(* IEC 61131-3 sources: trust-platform/examples/room_heating/libraries/plant/src, 22 files *)

(* ---- types.st ---- *)
(* The Plant library's shared types (specification trust-plant-library §3–§9). *)
NAMESPACE Plant

(* Who commands a device (§3): the program in Auto, the operator in Manual. *)
TYPE E_Mode : (Auto, Manual, OutOfService); END_TYPE

(* A measurement's quality (§7.1). *)
TYPE E_Quality : (Good, Uncertain, Bad); END_TYPE

(* A sequence's state (§9.4). *)
TYPE E_SequenceState : (Idle, Running, Held, Stopping, Stopped, Completed, Aborted, Failed); END_TYPE

END_NAMESPACE

(* ---- interfaces.st ---- *)
(* The capabilities of the Plant blocks (specification trust-plant-library §5). Each interface is
   small; a block implements the ones it supports. Operator commands return TRUE when accepted.
   An HMI button may call only a method of an interface its block implements. *)
NAMESPACE Plant

(* Mode and reset, common to every device (§3). *)
INTERFACE IDevice
    METHOD SetMode : BOOL
    VAR_INPUT
        Value : E_Mode;
    END_VAR
    END_METHOD
    METHOD GetMode : E_Mode
    END_METHOD
    METHOD Reset : BOOL
    END_METHOD
END_INTERFACE

INTERFACE IRunDevice EXTENDS IDevice
    METHOD Start : BOOL
    END_METHOD
    METHOD Stop : BOOL
    END_METHOD
    METHOD IsRunning : BOOL
    END_METHOD
END_INTERFACE

INTERFACE ISpeedDevice EXTENDS IRunDevice
    METHOD SetSpeed : BOOL
    VAR_INPUT
        Value : LREAL;
    END_VAR
    END_METHOD
END_INTERFACE

INTERFACE IPowerDevice EXTENDS IRunDevice
    METHOD SetPower : BOOL
    VAR_INPUT
        Value : LREAL;
    END_VAR
    END_METHOD
END_INTERFACE

INTERFACE IReversingDevice EXTENDS IDevice
    METHOD StartForward : BOOL
    END_METHOD
    METHOD StartReverse : BOOL
    END_METHOD
    METHOD Stop : BOOL
    END_METHOD
END_INTERFACE

INTERFACE ITwoSpeedDevice EXTENDS IDevice
    METHOD StartSlow : BOOL
    END_METHOD
    METHOD StartFast : BOOL
    END_METHOD
    METHOD Stop : BOOL
    END_METHOD
END_INTERFACE

INTERFACE IOpenCloseDevice EXTENDS IDevice
    METHOD Open : BOOL
    END_METHOD
    METHOD Close : BOOL
    END_METHOD
    METHOD IsOpen : BOOL
    END_METHOD
    METHOD IsClosed : BOOL
    END_METHOD
END_INTERFACE

(* A motor-operated valve can stop between its end positions. *)
INTERFACE ITravelStop
    METHOD StopTravel : BOOL
    END_METHOD
END_INTERFACE

INTERFACE IExtendRetractDevice EXTENDS IDevice
    METHOD Extend : BOOL
    END_METHOD
    METHOD Retract : BOOL
    END_METHOD
    METHOD IsExtended : BOOL
    END_METHOD
    METHOD IsRetracted : BOOL
    END_METHOD
END_INTERFACE

INTERFACE IPositionDevice EXTENDS IDevice
    METHOD SetPosition : BOOL
    VAR_INPUT
        Value : LREAL;
    END_VAR
    END_METHOD
    METHOD GetPosition : LREAL
    END_METHOD
END_INTERFACE

(* A device that a controller drives through its Auto value (§5): FollowsAuto is TRUE while the
   device follows that value now, GetActualValue is what the device does. A loop tracks
   GetActualValue while FollowsAuto is FALSE (§8.1), so it neither winds up nor bumps when the
   device follows it again. *)
INTERFACE IControlledDevice
    METHOD FollowsAuto : BOOL
    END_METHOD
    METHOD GetActualValue : LREAL
    END_METHOD
END_INTERFACE

(* An Engineer confirms that the service is done (§4.7). *)
INTERFACE IServiceable
    METHOD ServiceDone : BOOL
    END_METHOD
END_INTERFACE

(* A run device a group can command in Auto (§9.2). *)
INTERFACE IDutyMember EXTENDS IRunDevice
    METHOD IsAvailable : BOOL
    END_METHOD
    METHOD Demand
    VAR_INPUT
        Run : BOOL;
    END_VAR
    END_METHOD
    METHOD GetRunHours : LREAL
    END_METHOD
END_INTERFACE

INTERFACE IMeasurement
    METHOD GetValue : LREAL
    END_METHOD
    METHOD GetQuality : E_Quality
    END_METHOD
END_INTERFACE

INTERFACE ITotal
    METHOD ResetTotal : BOOL
    END_METHOD
END_INTERFACE

INTERFACE ICounter
    METHOD ResetCount : BOOL
    END_METHOD
END_INTERFACE

INTERFACE ITare
    METHOD Tare : BOOL
    END_METHOD
    METHOD ClearTare : BOOL
    END_METHOD
END_INTERFACE

INTERFACE ISetpoint
    METHOD SetSetpoint : BOOL
    VAR_INPUT
        Value : LREAL;
    END_VAR
    END_METHOD
END_INTERFACE

(* An Engineer bypasses one condition of a set for a limited time (§9.1). *)
INTERFACE IBypass
    METHOD Bypass : BOOL
    VAR_INPUT
        Index : INT;
    END_VAR
    END_METHOD
    METHOD RemoveBypass : BOOL
    VAR_INPUT
        Index : INT;
    END_VAR
    END_METHOD
END_INTERFACE

(* The alarms a block holds, for an alarm manager (§4.5, §9.3). *)
INTERFACE IAlarmSource
    METHOD GetAlarmCount : INT
    END_METHOD
    METHOD GetAlarm : REF_TO Alarm.Alarm
    VAR_INPUT
        Index : INT;
    END_VAR
    END_METHOD
END_INTERFACE

INTERFACE IAlarmManager
    METHOD AcknowledgeAll : BOOL
    END_METHOD
    METHOD Silence : BOOL
    END_METHOD
END_INTERFACE

INTERFACE ISequence
    METHOD Start : BOOL
    END_METHOD
    METHOD Stop : BOOL
    END_METHOD
    METHOD Hold : BOOL
    END_METHOD
    METHOD Resume : BOOL
    END_METHOD
    METHOD Abort : BOOL
    END_METHOD
    METHOD Reset : BOOL
    END_METHOD
    METHOD GetState : E_SequenceState
    END_METHOD
END_INTERFACE

INTERFACE ISequenceManager
    METHOD StopAll : BOOL
    END_METHOD
    METHOD AbortAll : BOOL
    END_METHOD
END_INTERFACE

END_NAMESPACE

(* ---- analog_input.st ---- *)
(* Analog instruments (specification trust-plant-library §7.1): scaling, quality, the optional
   Control.LowPass filter and four limit alarms. A broken signal raises one signal alarm and
   suppresses the limit alarms. The defaults suit a 4-20 mA signal (NAMUR NE 43); set RawLow,
   RawHigh, BadBelow and BadAbove for other signals. *)
NAMESPACE Plant
USING Alarm;
USING Control;

FUNCTION_BLOCK FB_AnalogInput IMPLEMENTS IMeasurement, IAlarmSource
VAR_INPUT
    (* The channel's value, for example in mA. *)
    Raw : LREAL;
    (* The I/O module's diagnosis for this channel. *)
    SignalFault : BOOL;
END_VAR
VAR PUBLIC
    Unit : STRING[16];
END_VAR
VAR PUBLIC RETAIN
    RawLow : LREAL := 4.0;
    RawHigh : LREAL := 20.0;
    RangeLow : LREAL := 0.0;
    RangeHigh : LREAL := 100.0;
    BadBelow : LREAL := 3.6;
    BadAbove : LREAL := 21.0;
    FilterTime : TIME := T#0s;
    HighHighEnabled : BOOL;
    HighEnabled : BOOL;
    LowEnabled : BOOL;
    LowLowEnabled : BOOL;
    HighHighLimit : LREAL := 95.0;
    HighLimit : LREAL := 90.0;
    LowLimit : LREAL := 10.0;
    LowLowLimit : LREAL := 5.0;
    Deadband : LREAL := 1.0;
    AlarmDelay : TIME := T#0s;
END_VAR
VAR_OUTPUT NON_RETAIN
    Value : LREAL;
    Percent : LREAL;
    Quality : E_Quality := E_Quality#Bad;
    Fault : BOOL;
    HighHigh : BOOL;
    High : BOOL;
    Low : BOOL;
    LowLow : BOOL;
END_VAR
VAR NON_RETAIN
    Filter : LowPass;
    Filtering : BOOL;
    HasValue : BOOL;
    Clock : FB_ScanClock;
    SignalAlarm : Alarm.DigitalAlarm;
    HighHighAlarm : Alarm.LimitAlarm;
    HighAlarm : Alarm.LimitAlarm;
    LowAlarm : Alarm.LimitAlarm;
    LowLowAlarm : Alarm.LimitAlarm;
END_VAR
    Measure();

METHOD PROTECTED Measure
VAR
    Span : LREAL;
    Range : LREAL;
    Scaled : LREAL;
    Parameters : LowPassParameters;
END_VAR
    Clock();
    Span := RawHigh - RawLow;
    Range := RangeHigh - RangeLow;
    IF NOT SignalFault AND F_Finite(Raw) AND Raw >= BadBelow AND Raw <= BadAbove
        AND F_Finite(Span) AND Span <> 0.0 THEN
        Scaled := RangeLow + (Raw - RawLow) * Range / Span;
        IF FilterTime > T#0s AND HasValue THEN
            Parameters.TimeConstant := F_Seconds(FilterTime);
            Parameters.Order := FilterOrder#FirstOrder;
            Filter.Configure(Parameters := Parameters);
            IF NOT Filtering THEN
                Filter.Initialize(Input := Value);
                Filtering := TRUE;
            END_IF;
            IF Clock.Seconds > 0.0 THEN
                Value := Filter.Update(Input := Scaled, CycleTime := Clock.Seconds);
            END_IF;
        ELSE
            Value := Scaled;
            Filtering := FALSE;
        END_IF;
        HasValue := TRUE;
        Quality := E_Quality#Good;
    ELSE
        (* The value holds its last good reading. *)
        Quality := E_Quality#Bad;
        Filtering := FALSE;
    END_IF;
    Fault := Quality = E_Quality#Bad;
    IF Range <> 0.0 AND F_Finite(Range) THEN
        Percent := (Value - RangeLow) / Range * 100.0;
    ELSE
        Percent := 0.0;
    END_IF;

    (* A limit that is not enabled, and every limit while the signal is bad, is suppressed: it
       does not annunciate and its output stays FALSE. *)
    SignalAlarm(Condition := Fault, Message := 'Signal fault', Priority := AlarmPriority#Medium);
    HighHighAlarm(Value := Value, Limit := HighHighLimit, Deadband := ABS(Deadband),
        Direction := LimitDirection#High, OnDelay := AlarmDelay, Suppressed := Fault OR NOT HighHighEnabled,
        Message := 'High-high', Priority := AlarmPriority#High);
    HighAlarm(Value := Value, Limit := HighLimit, Deadband := ABS(Deadband),
        Direction := LimitDirection#High, OnDelay := AlarmDelay, Suppressed := Fault OR NOT HighEnabled,
        Message := 'High', Priority := AlarmPriority#Medium);
    LowAlarm(Value := Value, Limit := LowLimit, Deadband := ABS(Deadband),
        Direction := LimitDirection#Low, OnDelay := AlarmDelay, Suppressed := Fault OR NOT LowEnabled,
        Message := 'Low', Priority := AlarmPriority#Medium);
    LowLowAlarm(Value := Value, Limit := LowLowLimit, Deadband := ABS(Deadband),
        Direction := LimitDirection#Low, OnDelay := AlarmDelay, Suppressed := Fault OR NOT LowLowEnabled,
        Message := 'Low-low', Priority := AlarmPriority#High);
    HighHigh := HighHighAlarm.Active AND NOT HighHighAlarm.SuppressedByDesign;
    High := HighAlarm.Active AND NOT HighAlarm.SuppressedByDesign;
    Low := LowAlarm.Active AND NOT LowAlarm.SuppressedByDesign;
    LowLow := LowLowAlarm.Active AND NOT LowLowAlarm.SuppressedByDesign;
END_METHOD

METHOD PUBLIC GetValue : LREAL
    GetValue := Value;
END_METHOD

METHOD PUBLIC GetQuality : E_Quality
    GetQuality := Quality;
END_METHOD

METHOD PUBLIC GetAlarmCount : INT
    GetAlarmCount := 5;
END_METHOD

METHOD PUBLIC GetAlarm : REF_TO Alarm.Alarm
VAR_INPUT
    Index : INT;
END_VAR
    CASE Index OF
        1: GetAlarm := REF(SignalAlarm);
        2: GetAlarm := REF(HighHighAlarm);
        3: GetAlarm := REF(HighAlarm);
        4: GetAlarm := REF(LowAlarm);
        5: GetAlarm := REF(LowLowAlarm);
    ELSE
        GetAlarm := NULL;
    END_CASE;
END_METHOD
END_FUNCTION_BLOCK

(* The instruments below differ in name and symbol; their unit comes from the instance. *)
FUNCTION_BLOCK FB_LevelInput EXTENDS FB_AnalogInput
    Measure();
END_FUNCTION_BLOCK

FUNCTION_BLOCK FB_PressureInput EXTENDS FB_AnalogInput
    Measure();
END_FUNCTION_BLOCK

FUNCTION_BLOCK FB_TemperatureInput EXTENDS FB_AnalogInput
    Measure();
END_FUNCTION_BLOCK

FUNCTION_BLOCK FB_AnalyzerInput EXTENDS FB_AnalogInput
    Measure();
END_FUNCTION_BLOCK

(* A flow instrument with its own totaliser on its measured value (§7.1.6). *)
FUNCTION_BLOCK FB_FlowInput EXTENDS FB_AnalogInput IMPLEMENTS ITotal
VAR_OUTPUT RETAIN
    (* Retained as well as the totaliser's, so it reads right before the first scan. *)
    Total : LREAL;
END_VAR
VAR PUBLIC RETAIN
    (* The time base of the flow's unit: T#1h for m3/h. *)
    TotalPer : TIME := T#1h;
END_VAR
VAR
    Totalizer : FB_Totalizer;
END_VAR
    Measure();
    Totalizer.TotalPer := TotalPer;
    Totalizer(Rate := Value, RateGood := Quality = E_Quality#Good);
    Total := Totalizer.Total;

METHOD PUBLIC ResetTotal : BOOL
    ResetTotal := Totalizer.ResetTotal();
    Total := 0.0;
END_METHOD
END_FUNCTION_BLOCK

END_NAMESPACE

(* ---- conditions.st ---- *)
(* Condition sets (specification trust-plant-library §9.1): up to eight conditions with texts, a
   first-out text, and Engineer bypasses that end by themselves. Interlocks and permissives may
   be bypassed; protection may not. These are ordinary process conditions, not certified safety
   functions. *)
NAMESPACE Plant

FUNCTION_BLOCK ABSTRACT FB_ConditionSet
VAR_INPUT
    (* TRUE while the condition is healthy; an unused condition stays TRUE. *)
    Condition1 : BOOL := TRUE;
    Condition2 : BOOL := TRUE;
    Condition3 : BOOL := TRUE;
    Condition4 : BOOL := TRUE;
    Condition5 : BOOL := TRUE;
    Condition6 : BOOL := TRUE;
    Condition7 : BOOL := TRUE;
    Condition8 : BOOL := TRUE;
    Text1 : STRING[80];
    Text2 : STRING[80];
    Text3 : STRING[80];
    Text4 : STRING[80];
    Text5 : STRING[80];
    Text6 : STRING[80];
    Text7 : STRING[80];
    Text8 : STRING[80];
END_VAR
VAR_OUTPUT NON_RETAIN
    (* Every condition healthy or bypassed. *)
    Healthy : BOOL := TRUE;
    Active : BOOL;
    (* The first condition that became unhealthy, held until all are healthy again. *)
    Text : STRING[80];
    FirstOut : INT;
    States : ARRAY[1..8] OF BOOL;
    Bypassed : ARRAY[1..8] OF BOOL;
    BypassActive : BOOL;
    (* The conditions a panel shows: each with a text, and any that is not healthy. *)
    InUse : ARRAY[1..8] OF BOOL;
END_VAR
VAR PUBLIC RETAIN
    BypassTime : TIME := T#1h;
END_VAR
VAR NON_RETAIN
    BypassTimers : ARRAY[1..8] OF TON;
END_VAR

METHOD PROTECTED Evaluate
VAR
    Texts : ARRAY[1..8] OF STRING[80];
    Index : INT;
    AllHealthy : BOOL;
    AnyBypass : BOOL;
END_VAR
    States[1] := Condition1;
    States[2] := Condition2;
    States[3] := Condition3;
    States[4] := Condition4;
    States[5] := Condition5;
    States[6] := Condition6;
    States[7] := Condition7;
    States[8] := Condition8;
    Texts[1] := Text1;
    Texts[2] := Text2;
    Texts[3] := Text3;
    Texts[4] := Text4;
    Texts[5] := Text5;
    Texts[6] := Text6;
    Texts[7] := Text7;
    Texts[8] := Text8;
    AllHealthy := TRUE;
    AnyBypass := FALSE;
    FOR Index := 1 TO 8 DO
        InUse[Index] := Texts[Index] <> '' OR NOT States[Index];
        BypassTimers[Index](IN := Bypassed[Index], PT := BypassTime);
        IF BypassTimers[Index].Q THEN
            Bypassed[Index] := FALSE;
            BypassTimers[Index](IN := FALSE, PT := BypassTime);
        END_IF;
        IF Bypassed[Index] THEN
            AnyBypass := TRUE;
        ELSIF NOT States[Index] THEN
            AllHealthy := FALSE;
            IF FirstOut = 0 THEN
                FirstOut := Index;
            END_IF;
        END_IF;
    END_FOR;
    IF AllHealthy THEN
        FirstOut := 0;
    END_IF;
    Healthy := AllHealthy;
    Active := NOT AllHealthy;
    BypassActive := AnyBypass;
    IF FirstOut = 0 THEN
        Text := '';
    ELSIF Texts[FirstOut] = '' THEN
        Text := CONCAT('Condition ', INT_TO_STRING(FirstOut));
    ELSE
        Text := Texts[FirstOut];
    END_IF;
END_METHOD

(* Bypass one condition for BypassTime; a repeated bypass restarts the time. *)
METHOD PROTECTED BypassCondition : BOOL
VAR_INPUT
    Index : INT;
END_VAR
    BypassCondition := Index >= 1 AND Index <= 8;
    IF BypassCondition THEN
        Bypassed[Index] := TRUE;
        BypassTimers[Index](IN := FALSE, PT := BypassTime);
    END_IF;
END_METHOD

METHOD PROTECTED EndBypass : BOOL
VAR_INPUT
    Index : INT;
END_VAR
    EndBypass := Index >= 1 AND Index <= 8;
    IF EndBypass THEN
        Bypassed[Index] := FALSE;
    END_IF;
END_METHOD
END_FUNCTION_BLOCK

(* Interlocks: wire Active and Text to a device's Interlock and InterlockText. *)
FUNCTION_BLOCK FB_Interlocks EXTENDS FB_ConditionSet IMPLEMENTS IBypass
    Evaluate();

METHOD PUBLIC Bypass : BOOL
VAR_INPUT
    Index : INT;
END_VAR
    Bypass := BypassCondition(Index := Index);
END_METHOD

METHOD PUBLIC RemoveBypass : BOOL
VAR_INPUT
    Index : INT;
END_VAR
    RemoveBypass := EndBypass(Index := Index);
END_METHOD
END_FUNCTION_BLOCK

(* Permissives: wire Healthy and Text to a device's Permissive and PermissiveText. *)
FUNCTION_BLOCK FB_Permissives EXTENDS FB_ConditionSet IMPLEMENTS IBypass
    Evaluate();

METHOD PUBLIC Bypass : BOOL
VAR_INPUT
    Index : INT;
END_VAR
    Bypass := BypassCondition(Index := Index);
END_METHOD

METHOD PUBLIC RemoveBypass : BOOL
VAR_INPUT
    Index : INT;
END_VAR
    RemoveBypass := EndBypass(Index := Index);
END_METHOD
END_FUNCTION_BLOCK

(* Equipment protection: like interlocks, without bypass. *)
FUNCTION_BLOCK FB_Protection EXTENDS FB_ConditionSet
    Evaluate();
END_FUNCTION_BLOCK

END_NAMESPACE

(* ---- control_valve.st ---- *)
(* Control valves and modulating dampers (specification trust-plant-library §6.9). The safe state
   is FailPosition. Leaving it is a start: it needs the permissive; once released the valve keeps
   following its position when the permissive drops. *)
NAMESPACE Plant
USING Alarm;

FUNCTION_BLOCK FB_ControlValve EXTENDS FB_Device IMPLEMENTS IPositionDevice, IAlarmSource, IControlledDevice
VAR_INPUT
    (* The program's position in % open, followed in Auto. *)
    AutoPosition : LREAL;
    PositionFeedback : LREAL;
    HasFeedback : BOOL;
    (* The position the valve takes on loss of signal or air, in % open. *)
    FailPosition : LREAL;
END_VAR
VAR_OUTPUT NON_RETAIN
    (* The positioner's setpoint in % open. *)
    PositionSetpoint : LREAL;
    Position : LREAL;
    InPosition : BOOL;
    (* The operator's position in % open. *)
    ManualPosition : LREAL;
    Deviating : BOOL;
END_VAR
VAR PUBLIC RETAIN
    MinPosition : LREAL := 0.0;
    MaxPosition : LREAL := 100.0;
    PositionDeviation : LREAL := 5.0;
    DeviationTime : TIME := T#10s;
END_VAR
VAR NON_RETAIN
    Released : BOOL;
    Initialized : BOOL;
    DeviationAlarm : Alarm.DigitalAlarm;
END_VAR
    ExecutePosition();

METHOD PROTECTED ExecutePosition
VAR
    Low : LREAL;
    High : LREAL;
    Wanted : LREAL;
    Supervised : BOOL;
END_VAR
    (* After a restart a manually positioned valve is at its fail position (§4.8). *)
    IF NOT Initialized THEN
        ManualPosition := FailPosition;
        PositionSetpoint := FailPosition;
        Initialized := TRUE;
    END_IF;
    (* A control valve latches no fault, so a Reset has nothing to clear. *)
    ResetRequested := FALSE;
    Supervised := Mode <> E_Mode#OutOfService;
    Low := MIN(MinPosition, MaxPosition);
    High := MAX(MinPosition, MaxPosition);
    Fault := FALSE;
    FaultText := '';
    IF HeldSafe() THEN
        Released := FALSE;
    ELSIF NOT Released AND MayStart() THEN
        Released := TRUE;
    END_IF;
    IF Mode = E_Mode#Auto THEN
        Wanted := AutoPosition;
        IF NOT F_Finite(Wanted) THEN
            Wanted := PositionSetpoint;
        END_IF;
    ELSE
        Wanted := ManualPosition;
    END_IF;
    IF Released THEN
        PositionSetpoint := LIMIT(Low, Wanted, High);
    ELSE
        PositionSetpoint := FailPosition;
    END_IF;
    IF HasFeedback THEN
        Position := PositionFeedback;
    ELSE
        Position := PositionSetpoint;
    END_IF;
    Deviating := HasFeedback AND Supervised
        AND (NOT F_Finite(PositionFeedback) OR ABS(PositionFeedback - PositionSetpoint) > PositionDeviation);
    InPosition := NOT Deviating;
    (* Bumpless (§3.4): Manual holds the valve where it is; the safe state leaves it at the fail
       position. *)
    ManualPosition := PositionSetpoint;
    DeviationAlarm(Condition := Deviating, OnDelay := DeviationTime, Suppressed := NOT Supervised,
        Message := 'Position deviation', Priority := AlarmPriority#Low);
    Publish();
END_METHOD

(* Accepted in Manual while nothing blocks the valve; clamped to MinPosition..MaxPosition. *)
METHOD PUBLIC SetPosition : BOOL
VAR_INPUT
    Value : LREAL;
END_VAR
    SetPosition := AcceptsStart() AND F_Finite(Value);
    IF SetPosition THEN
        ManualPosition := LIMIT(MIN(MinPosition, MaxPosition), Value, MAX(MinPosition, MaxPosition));
    END_IF;
END_METHOD

METHOD PUBLIC GetPosition : LREAL
    GetPosition := Position;
END_METHOD

METHOD PUBLIC GetAlarmCount : INT
    GetAlarmCount := 1;
END_METHOD

METHOD PUBLIC GetAlarm : REF_TO Alarm.Alarm
VAR_INPUT
    Index : INT;
END_VAR
    IF Index = 1 THEN
        GetAlarm := REF(DeviationAlarm);
    ELSE
        GetAlarm := NULL;
    END_IF;
END_METHOD

(* The valve follows its Auto position while in Auto and released from its fail position
   (§6.9); a controller that drives it tracks Position otherwise (§8.1). *)
METHOD PUBLIC FollowsAuto : BOOL
    FollowsAuto := Mode = E_Mode#Auto AND Released;
END_METHOD

METHOD PUBLIC GetActualValue : LREAL
    GetActualValue := Position;
END_METHOD

END_FUNCTION_BLOCK

FUNCTION_BLOCK FB_ModulatingDamper EXTENDS FB_ControlValve
    ExecutePosition();
END_FUNCTION_BLOCK

END_NAMESPACE

(* ---- controllers.st ---- *)
(* Controllers (specification trust-plant-library §8). A PID loop is no block of this library: Create
   PLC code writes it as ordinary code around the Control library's PID (specification 39, §10.5).
   The thermostat-style on/off controller is a block. *)
NAMESPACE Plant

(* A thermostat-style controller (§8.3): Demand is TRUE below the setpoint for heating (above it
   for cooling), with Hysteresis around the setpoint. Wire Demand to a device's Auto input. *)
FUNCTION_BLOCK FB_OnOffController IMPLEMENTS ISetpoint
VAR_INPUT
    (* The measured value: an instrument by composition, else ProcessValue and its quality. *)
    Measurement : IMeasurement;
    ProcessValue : LREAL;
    ProcessValueGood : BOOL := TRUE;
END_VAR
VAR_OUTPUT RETAIN
    Setpoint : LREAL := 50.0;
END_VAR
VAR_OUTPUT NON_RETAIN
    Demand : BOOL;
    MeasuredValue : LREAL;
END_VAR
VAR PUBLIC RETAIN
    Hysteresis : LREAL := 1.0;
    (* TRUE: demand below the setpoint; FALSE (cooling): demand above it. *)
    Heating : BOOL := TRUE;
    SetpointMin : LREAL := 0.0;
    SetpointMax : LREAL := 100.0;
END_VAR
VAR_TEMP
    Half : LREAL;
    Measured : LREAL;
    Good : BOOL;
END_VAR
    Half := ABS(Hysteresis) / 2.0;
    IF Measurement <> NULL THEN
        Measured := Measurement.GetValue();
        Good := Measurement.GetQuality() = E_Quality#Good;
    ELSE
        Measured := ProcessValue;
        Good := ProcessValueGood;
    END_IF;
    IF Good AND F_Finite(Measured) THEN
        MeasuredValue := Measured;
    END_IF;
    IF NOT Good OR NOT F_Finite(Measured) THEN
        Demand := FALSE;
    ELSIF Heating THEN
        IF Measured < Setpoint - Half THEN
            Demand := TRUE;
        ELSIF Measured > Setpoint + Half THEN
            Demand := FALSE;
        END_IF;
    ELSE
        IF Measured > Setpoint + Half THEN
            Demand := TRUE;
        ELSIF Measured < Setpoint - Half THEN
            Demand := FALSE;
        END_IF;
    END_IF;

METHOD PUBLIC SetSetpoint : BOOL
VAR_INPUT
    Value : LREAL;
END_VAR
    SetSetpoint := F_Finite(Value);
    IF SetSetpoint THEN
        Setpoint := LIMIT(MIN(SetpointMin, SetpointMax), Value, MAX(SetpointMin, SetpointMax));
    END_IF;
END_METHOD
END_FUNCTION_BLOCK

END_NAMESPACE

(* ---- cylinder.st ---- *)
(* A pneumatic or hydraulic cylinder (specification trust-plant-library §6.8). Single-acting: one
   solenoid extends it and the spring retracts it, so the safe state is retracted. Double-acting:
   one solenoid each way; the safe state de-energises both and it stays where it is. *)
NAMESPACE Plant
USING Alarm;

FUNCTION_BLOCK FB_Cylinder EXTENDS FB_Device IMPLEMENTS IExtendRetractDevice, IAlarmSource
VAR_INPUT
    (* The program's position, followed in Auto: TRUE extended. *)
    AutoExtend : BOOL;
    ExtendedSensor : BOOL;
    RetractedSensor : BOOL;
    HasExtendedSensor : BOOL := TRUE;
    HasRetractedSensor : BOOL := TRUE;
    DoubleActing : BOOL;
END_VAR
VAR_OUTPUT NON_RETAIN
    (* Solenoid A, extending. *)
    ExtendCommand : BOOL;
    (* Solenoid B, retracting; double-acting only. *)
    RetractCommand : BOOL;
    Extended : BOOL;
    Retracted : BOOL;
    Moving : BOOL;
    FailedToExtend : BOOL;
    FailedToRetract : BOOL;
    FeedbackConflict : BOOL;
    ExtendPermit : BOOL;
    RetractPermit : BOOL;
END_VAR
VAR_OUTPUT RETAIN
    Operations : UDINT;
END_VAR
VAR PUBLIC RETAIN
    ExtendTimeout : TIME := T#5s;
    RetractTimeout : TIME := T#5s;
END_VAR
VAR NON_RETAIN
    (* The commanded position: TRUE extended. *)
    Wanted : BOOL;
    ManualExtend : BOOL;
    Watch : FB_EndPositionWatch;
    FailedToExtendAlarm : Alarm.DigitalAlarm;
    FailedToRetractAlarm : Alarm.DigitalAlarm;
    ConflictAlarm : Alarm.DigitalAlarm;
END_VAR
    ExecuteCylinder();

METHOD PROTECTED ExecuteCylinder
VAR
    Supervised : BOOL;
    Safe : BOOL;
    Desired : BOOL;
END_VAR
    Supervised := Mode <> E_Mode#OutOfService;
    CASE Mode OF
        E_Mode#Auto:
            Desired := AutoExtend;
        E_Mode#Manual:
            Desired := ManualExtend;
    ELSE
        Desired := FALSE;
    END_CASE;
    (* Extending, and with double action any movement, counts as a start. *)
    IF Desired <> Wanted AND (Desired OR DoubleActing) AND NOT MayStart() THEN
        Desired := Wanted;
    END_IF;
    Safe := HeldSafe();
    IF Safe AND NOT DoubleActing THEN
        Desired := FALSE;
    END_IF;
    Wanted := Desired;

    Watch(Enable := Supervised AND NOT (Safe AND DoubleActing), TowardsA := Wanted,
        AtA := ExtendedSensor, AtB := RetractedSensor, HasA := HasExtendedSensor,
        HasB := HasRetractedSensor, TimeoutA := ExtendTimeout, TimeoutB := RetractTimeout,
        Clear := TakeReset());
    FailedToExtend := Watch.FailedA;
    FailedToRetract := Watch.FailedB;
    FeedbackConflict := Watch.Conflict;
    Fault := FailedToExtend OR FailedToRetract OR FeedbackConflict;
    Safe := Safe OR Fault;
    IF Safe AND NOT DoubleActing THEN
        Wanted := FALSE;
    END_IF;
    IF Safe AND DoubleActing THEN
        ExtendCommand := FALSE;
        RetractCommand := FALSE;
    ELSE
        ExtendCommand := Wanted;
        RetractCommand := DoubleActing AND NOT Wanted;
    END_IF;
    Extended := Watch.InA;
    Retracted := Watch.InB;
    Moving := Watch.Moving AND NOT (Safe AND DoubleActing);
    IF FeedbackConflict THEN
        FaultText := 'Both end sensors active: check them, then reset';
    ELSIF FailedToExtend THEN
        FaultText := 'Failed to extend: reset to try again';
    ELSIF FailedToRetract THEN
        FaultText := 'Failed to retract: reset to try again';
    ELSE
        FaultText := '';
    END_IF;

    (* Bumpless (§3.4). *)
    ManualExtend := Wanted;

    FailedToExtendAlarm(Condition := FailedToExtend, Suppressed := NOT Supervised,
        Message := 'Failed to extend', Priority := AlarmPriority#Medium);
    FailedToRetractAlarm(Condition := FailedToRetract, Suppressed := NOT Supervised,
        Message := 'Failed to retract', Priority := AlarmPriority#Medium);
    ConflictAlarm(Condition := FeedbackConflict, Suppressed := NOT Supervised,
        Message := 'End sensors conflict', Priority := AlarmPriority#Medium);
    IF Supervised AND Watch.Arrived AND Operations < UDINT#4294967295 THEN
        Operations := Operations + 1;
    END_IF;
    Publish();
    ExtendPermit := StartPermit;
    RetractPermit := Manual AND (NOT DoubleActing OR NOT Blocked);
END_METHOD

METHOD PUBLIC Extend : BOOL
    Extend := AcceptsStart();
    IF Extend THEN
        ManualExtend := TRUE;
    END_IF;
END_METHOD

METHOD PUBLIC Retract : BOOL
    IF DoubleActing THEN
        Retract := AcceptsStart();
    ELSE
        Retract := AcceptsCommands();
    END_IF;
    IF Retract THEN
        ManualExtend := FALSE;
    END_IF;
END_METHOD

METHOD PUBLIC IsExtended : BOOL
    IsExtended := Extended;
END_METHOD

METHOD PUBLIC IsRetracted : BOOL
    IsRetracted := Retracted;
END_METHOD

METHOD PUBLIC GetAlarmCount : INT
    GetAlarmCount := 3;
END_METHOD

METHOD PUBLIC GetAlarm : REF_TO Alarm.Alarm
VAR_INPUT
    Index : INT;
END_VAR
    CASE Index OF
        1: GetAlarm := REF(FailedToExtendAlarm);
        2: GetAlarm := REF(FailedToRetractAlarm);
        3: GetAlarm := REF(ConflictAlarm);
    ELSE
        GetAlarm := NULL;
    END_CASE;
END_METHOD
END_FUNCTION_BLOCK

END_NAMESPACE

(* ---- device.st ---- *)
(* What every actuator shares (specification trust-plant-library §3, §4): the mode, the interlock
   and permissive, the latched fault and its reset, and the permits and texts the operator panels
   show. A concrete device takes the reset with TakeReset at the start of its scan, sets Fault and
   FaultText, and calls Publish at the end. *)
NAMESPACE Plant

FUNCTION_BLOCK ABSTRACT FB_Device IMPLEMENTS IDevice
VAR_INPUT
    (* While TRUE the device is held in its safe state in every mode. *)
    Interlock : BOOL;
    InterlockText : STRING[80];
    (* While FALSE a start is refused; a running device continues. *)
    Permissive : BOOL := TRUE;
    PermissiveText : STRING[80];
END_VAR
VAR_OUTPUT RETAIN
    Mode : E_Mode;
END_VAR
VAR_OUTPUT NON_RETAIN
    Manual : BOOL;
    OutOfService : BOOL;
    InService : BOOL := TRUE;
    (* A latched trip or supervision failure; Reset clears it once the cause is gone. *)
    Fault : BOOL;
    Interlocked : BOOL;
    (* A start would be refused now, and why. *)
    Blocked : BOOL;
    BlockReason : STRING[80];
    (* The operator may start the device now: Manual and not blocked. *)
    StartPermit : BOOL;
    (* Why an operator command is refused now; empty when it is accepted. *)
    CommandText : STRING[80];
    (* The panel's message line: why the device is blocked, else why a command is refused. *)
    ReasonText : STRING[80];
END_VAR
VAR NON_RETAIN
    ResetRequested : BOOL;
    FaultText : STRING[80];
END_VAR

METHOD PUBLIC SetMode : BOOL
VAR_INPUT
    Value : E_Mode;
END_VAR
    Mode := Value;
    UpdateMode();
    SetMode := TRUE;
END_METHOD

METHOD PUBLIC GetMode : E_Mode
    GetMode := Mode;
END_METHOD

(* Accepted in every mode; applied at the device's next scan. It never starts anything. *)
METHOD PUBLIC Reset : BOOL
    ResetRequested := TRUE;
    Reset := TRUE;
END_METHOD

(* TRUE once per Reset, at the start of the device's next scan. *)
METHOD PROTECTED TakeReset : BOOL
    TakeReset := ResetRequested;
    ResetRequested := FALSE;
END_METHOD

(* Nothing prevents a start: in service, no fault, no interlock and the permissive present. *)
METHOD PROTECTED MayStart : BOOL
    MayStart := Mode <> E_Mode#OutOfService AND NOT Fault AND NOT Interlock AND Permissive;
END_METHOD

(* An operator command applies only in Manual (§3.5). *)
METHOD PROTECTED AcceptsCommands : BOOL
    AcceptsCommands := Mode = E_Mode#Manual;
END_METHOD

(* An operator start applies in Manual while nothing blocks it. *)
METHOD PROTECTED AcceptsStart : BOOL
    AcceptsStart := Mode = E_Mode#Manual AND MayStart();
END_METHOD

(* The device is held in its safe state (§4.6). *)
METHOD PROTECTED HeldSafe : BOOL
    HeldSafe := Interlock OR Fault OR Mode = E_Mode#OutOfService;
END_METHOD

METHOD PROTECTED UpdateMode
    Manual := Mode = E_Mode#Manual;
    OutOfService := Mode = E_Mode#OutOfService;
    InService := NOT OutOfService;
END_METHOD

(* The state, the permits and the texts (§4.2), once Fault and FaultText are set for this scan. *)
METHOD PROTECTED Publish
    UpdateMode();
    Interlocked := Interlock;
    Blocked := OutOfService OR Fault OR Interlock OR NOT Permissive;
    IF OutOfService THEN
        BlockReason := 'Out of service';
    ELSIF Fault THEN
        BlockReason := FaultText;
    ELSIF Interlock THEN
        IF InterlockText = '' THEN
            BlockReason := 'Interlocked';
        ELSE
            BlockReason := CONCAT('Interlocked: ', InterlockText);
        END_IF;
    ELSIF NOT Permissive THEN
        IF PermissiveText = '' THEN
            BlockReason := 'Not permitted';
        ELSE
            BlockReason := CONCAT('Not permitted: ', PermissiveText);
        END_IF;
    ELSE
        BlockReason := '';
    END_IF;
    StartPermit := Manual AND NOT Blocked;
    IF Mode = E_Mode#Auto THEN
        CommandText := 'Auto: switch to Manual';
    ELSIF OutOfService THEN
        CommandText := 'Out of service';
    ELSIF Blocked THEN
        CommandText := BlockReason;
    ELSE
        CommandText := '';
    END_IF;
    IF BlockReason <> '' THEN
        ReasonText := BlockReason;
    ELSE
        ReasonText := CommandText;
    END_IF;
END_METHOD
END_FUNCTION_BLOCK

END_NAMESPACE

(* ---- digital_input.st ---- *)
(* Digital instruments (specification trust-plant-library §7.2): inversion, debounce, quality and
   an optional switch alarm. *)
NAMESPACE Plant
USING Alarm;

FUNCTION_BLOCK FB_DigitalInput IMPLEMENTS IAlarmSource
VAR_INPUT
    Input : BOOL;
    (* The I/O module's diagnosis for this channel. *)
    SignalFault : BOOL;
END_VAR
VAR PUBLIC RETAIN
    Invert : BOOL;
    Debounce : TIME := T#0s;
    AlarmEnabled : BOOL;
    (* The value that raises the switch alarm. *)
    AlarmWhen : BOOL := TRUE;
    AlarmText : STRING[80] := 'Switch active';
END_VAR
VAR_OUTPUT NON_RETAIN
    Value : BOOL;
    Quality : E_Quality := E_Quality#Bad;
END_VAR
VAR NON_RETAIN
    Initialized : BOOL;
    OnTimer : TON;
    OffTimer : TON;
    SwitchAlarm : Alarm.DigitalAlarm;
    SignalAlarm : Alarm.DigitalAlarm;
END_VAR
    Sense();

METHOD PROTECTED Sense
VAR
    Level : BOOL;
END_VAR
    Level := Input XOR Invert;
    IF NOT Initialized THEN
        Value := Level;
        Initialized := TRUE;
    END_IF;
    OnTimer(IN := Level AND NOT Value, PT := Debounce);
    OffTimer(IN := NOT Level AND Value, PT := Debounce);
    IF OnTimer.Q THEN
        Value := TRUE;
    ELSIF OffTimer.Q THEN
        Value := FALSE;
    END_IF;
    IF SignalFault THEN
        Quality := E_Quality#Bad;
    ELSE
        Quality := E_Quality#Good;
    END_IF;
    SwitchAlarm(Condition := AlarmEnabled AND Value = AlarmWhen, Suppressed := SignalFault,
        Message := AlarmText, Priority := AlarmPriority#Medium);
    SignalAlarm(Condition := SignalFault, Message := 'Signal fault', Priority := AlarmPriority#Medium);
END_METHOD

METHOD PUBLIC GetAlarmCount : INT
    GetAlarmCount := 2;
END_METHOD

METHOD PUBLIC GetAlarm : REF_TO Alarm.Alarm
VAR_INPUT
    Index : INT;
END_VAR
    CASE Index OF
        1: GetAlarm := REF(SwitchAlarm);
        2: GetAlarm := REF(SignalAlarm);
    ELSE
        GetAlarm := NULL;
    END_CASE;
END_METHOD
END_FUNCTION_BLOCK

FUNCTION_BLOCK FB_LevelSwitch EXTENDS FB_DigitalInput
    Sense();
END_FUNCTION_BLOCK

FUNCTION_BLOCK FB_PressureSwitch EXTENDS FB_DigitalInput
    Sense();
END_FUNCTION_BLOCK

END_NAMESPACE

(* ---- drive.st ---- *)
(* Variable-speed motors (specification trust-plant-library §6.2): run control from FB_RunDevice
   plus a speed reference for the drive. A drive starts at 0 %: the operator's speed is 0 % after
   a restart and after every stop. *)
NAMESPACE Plant
USING Alarm;

FUNCTION_BLOCK FB_VariableSpeedMotor EXTENDS FB_RunDevice IMPLEMENTS ISpeedDevice, IControlledDevice
VAR_INPUT
    (* The program's speed in %, followed in Auto while running. *)
    AutoSpeed : LREAL;
    SpeedFeedback : LREAL;
    HasSpeedFeedback : BOOL;
END_VAR
VAR_OUTPUT NON_RETAIN
    (* The drive's speed reference in %. *)
    SpeedSetpoint : LREAL;
    Speed : LREAL;
    (* The operator's speed in %. *)
    ManualSpeed : LREAL;
    SpeedDeviating : BOOL;
END_VAR
VAR PUBLIC RETAIN
    MinSpeed : LREAL := 0.0;
    MaxSpeed : LREAL := 100.0;
    SpeedDeviation : LREAL := 5.0;
    DeviationTime : TIME := T#10s;
END_VAR
VAR NON_RETAIN
    WasCommanded : BOOL;
    SpeedDeviationAlarm : Alarm.DigitalAlarm;
END_VAR
    ExecuteRun();
    ExecuteSpeed();

METHOD PROTECTED ExecuteSpeed
VAR
    Low : LREAL;
    High : LREAL;
    Wanted : LREAL;
END_VAR
    Low := MIN(MinSpeed, MaxSpeed);
    High := MAX(MinSpeed, MaxSpeed);
    IF RunCommand THEN
        IF Mode = E_Mode#Auto THEN
            Wanted := AutoSpeed;
            IF NOT F_Finite(Wanted) THEN
                Wanted := SpeedSetpoint;
            END_IF;
            (* Bumpless: Manual continues at the speed Auto had. *)
            ManualSpeed := LIMIT(Low, Wanted, High);
        ELSE
            Wanted := ManualSpeed;
        END_IF;
        SpeedSetpoint := LIMIT(Low, Wanted, High);
    ELSE
        SpeedSetpoint := 0.0;
        IF WasCommanded THEN
            ManualSpeed := 0.0;
        END_IF;
    END_IF;
    WasCommanded := RunCommand;
    IF HasSpeedFeedback THEN
        Speed := SpeedFeedback;
    ELSE
        Speed := SpeedSetpoint;
    END_IF;
    SpeedDeviating := HasSpeedFeedback AND RunCommand
        AND (NOT F_Finite(SpeedFeedback) OR ABS(SpeedFeedback - SpeedSetpoint) > SpeedDeviation);
    SpeedDeviationAlarm(Condition := SpeedDeviating, OnDelay := DeviationTime,
        Suppressed := Mode = E_Mode#OutOfService, Message := 'Speed deviation', Priority := AlarmPriority#Low);
END_METHOD

(* Accepted in Manual, also while stopped, so a speed can be chosen before the start. *)
METHOD PUBLIC SetSpeed : BOOL
VAR_INPUT
    Value : LREAL;
END_VAR
    SetSpeed := AcceptsCommands() AND F_Finite(Value);
    IF SetSpeed THEN
        ManualSpeed := LIMIT(MIN(MinSpeed, MaxSpeed), Value, MAX(MinSpeed, MaxSpeed));
    END_IF;
END_METHOD

METHOD PUBLIC OVERRIDE GetAlarmCount : INT
    GetAlarmCount := 4;
END_METHOD

METHOD PUBLIC OVERRIDE GetAlarm : REF_TO Alarm.Alarm
VAR_INPUT
    Index : INT;
END_VAR
    IF Index = 4 THEN
        GetAlarm := REF(SpeedDeviationAlarm);
    ELSE
        GetAlarm := SUPER.GetAlarm(Index);
    END_IF;
END_METHOD

(* The drive follows its Auto speed while in Auto and running (§6.2); a controller that drives it
   tracks Speed otherwise (§8.1). *)
METHOD PUBLIC FollowsAuto : BOOL
    FollowsAuto := Mode = E_Mode#Auto AND RunCommand;
END_METHOD

METHOD PUBLIC GetActualValue : LREAL
    GetActualValue := Speed;
END_METHOD

END_FUNCTION_BLOCK

FUNCTION_BLOCK FB_VariableSpeedPump EXTENDS FB_VariableSpeedMotor
    ExecuteRun();
    ExecuteSpeed();
END_FUNCTION_BLOCK

FUNCTION_BLOCK FB_VariableSpeedFan EXTENDS FB_VariableSpeedMotor
    ExecuteRun();
    ExecuteSpeed();
END_FUNCTION_BLOCK

FUNCTION_BLOCK FB_DosingPump EXTENDS FB_VariableSpeedMotor
    ExecuteRun();
    ExecuteSpeed();
END_FUNCTION_BLOCK

END_NAMESPACE

(* ---- end_position.st ---- *)
(* Supervision of a two-position actuator (specification trust-plant-library §6.6–§6.8), shared by
   the on/off valve, the damper and the cylinder. Position A is open or extended, B closed or
   retracted. Without a switch, that end position follows the command. *)
NAMESPACE Plant

FUNCTION_BLOCK FB_EndPositionWatch
VAR_INPUT
    (* FALSE out of service, or while nothing is commanded. *)
    Enable : BOOL;
    (* Commanded to A; else to B. *)
    TowardsA : BOOL;
    AtA : BOOL;
    AtB : BOOL;
    HasA : BOOL;
    HasB : BOOL;
    TimeoutA : TIME;
    TimeoutB : TIME;
    (* A reset: clears the latched failures and restarts the timing. *)
    Clear : BOOL;
END_VAR
VAR_OUTPUT NON_RETAIN
    InA : BOOL;
    InB : BOOL;
    Moving : BOOL;
    FailedA : BOOL;
    FailedB : BOOL;
    Conflict : BOOL;
    (* TRUE for one scan when the commanded end position is reached: one operation. *)
    Arrived : BOOL;
END_VAR
VAR NON_RETAIN
    WatchA : TON;
    WatchB : TON;
    ConflictWatch : TON;
    WasInA : BOOL;
    WasInB : BOOL;
    Primed : BOOL;
END_VAR
    IF Clear THEN
        FailedA := FALSE;
        FailedB := FALSE;
        Conflict := FALSE;
        WatchA(IN := FALSE);
        WatchB(IN := FALSE);
        ConflictWatch(IN := FALSE);
    END_IF;
    IF HasA THEN
        InA := AtA;
    ELSE
        InA := TowardsA;
    END_IF;
    IF HasB THEN
        InB := AtB;
    ELSE
        InB := NOT TowardsA;
    END_IF;
    Moving := (TowardsA AND NOT InA) OR (NOT TowardsA AND NOT InB);
    (* Not reaching the commanded end position in time, or leaving it, is a failure. *)
    WatchA(IN := Enable AND TowardsA AND NOT InA, PT := TimeoutA);
    WatchB(IN := Enable AND NOT TowardsA AND NOT InB, PT := TimeoutB);
    ConflictWatch(IN := Enable AND HasA AND HasB AND AtA AND AtB, PT := T#1s);
    IF WatchA.Q THEN
        FailedA := TRUE;
    END_IF;
    IF WatchB.Q THEN
        FailedB := TRUE;
    END_IF;
    IF ConflictWatch.Q THEN
        Conflict := TRUE;
    END_IF;
    Arrived := Primed AND ((TowardsA AND InA AND NOT WasInA) OR (NOT TowardsA AND InB AND NOT WasInB));
    WasInA := InA;
    WasInB := InB;
    Primed := TRUE;
END_FUNCTION_BLOCK

END_NAMESPACE

(* ---- functions.st ---- *)
(* Small calculations shared by the blocks. *)
NAMESPACE Plant

(* TRUE for a finite number: neither NaN nor infinite. *)
FUNCTION F_Finite : BOOL
VAR_INPUT
    Value : LREAL;
END_VAR
    F_Finite := Value = Value AND ABS(Value) <= 1.7976931348623157E308;
END_FUNCTION

(* A duration in seconds. A negative duration counts as zero; durations are capped at 49 days,
   the range of the millisecond conversion. *)
FUNCTION F_Seconds : LREAL
VAR_INPUT
    Value : TIME;
END_VAR
    IF Value <= T#0s THEN
        F_Seconds := 0.0;
    ELSIF Value >= T#49d THEN
        F_Seconds := 4233600.0;
    ELSE
        F_Seconds := UDINT_TO_LREAL(DWORD_TO_UDINT(TIME_TO_DWORD(Value))) / 1000.0;
    END_IF;
END_FUNCTION

(* The time since the previous call, from the runtime clock; zero at the first call after a
   restart, so a restart never counts the time the PLC was off. *)
FUNCTION_BLOCK FB_ScanClock
VAR_OUTPUT
    Elapsed : TIME;
    Seconds : LREAL;
END_VAR
VAR NON_RETAIN
    Started : BOOL;
    Last : TIME;
END_VAR
VAR_TEMP
    Now : TIME;
END_VAR
    Now := TIME();
    IF Started AND Now >= Last THEN
        Elapsed := Now - Last;
    ELSE
        Elapsed := T#0s;
    END_IF;
    Started := TRUE;
    Last := Now;
    Seconds := F_Seconds(Elapsed);
END_FUNCTION_BLOCK

END_NAMESPACE

(* ---- groups.st ---- *)
(* Groups of interchangeable run devices (specification trust-plant-library §9.2). Members are
   chosen by composition: Member1..Member4 in the call. A group never registers anything; it
   commands its members through IDutyMember.Demand, which they follow only in Auto, and every
   member keeps its own interlocks, faults and supervision. *)
NAMESPACE Plant
USING Alarm;

FUNCTION_BLOCK ABSTRACT FB_Group IMPLEMENTS IAlarmSource
VAR_INPUT
    Member1 : IDutyMember;
    Member2 : IDutyMember;
    Member3 : IDutyMember;
    Member4 : IDutyMember;
END_VAR
VAR_OUTPUT NON_RETAIN
    (* How many members run, are available, and the group wants running. *)
    RunningCount : INT;
    AvailableCount : INT;
    Target : INT;
    (* Fewer members run than wanted, for longer than ShortfallDelay. *)
    Shortfall : BOOL;
    Selected : ARRAY[1..4] OF BOOL;
END_VAR
VAR PUBLIC RETAIN
    (* The member to start first when available; 0 chooses by fewest run hours. *)
    Preferred : INT := 0;
    StartDelay : TIME := T#2s;
    StopDelay : TIME := T#2s;
    ShortfallDelay : TIME := T#10s;
END_VAR
VAR NON_RETAIN
    Members : ARRAY[1..4] OF IDutyMember;
    Changed : BOOL;
    SinceChange : TON;
    ShortfallTimer : TON;
    ShortfallAlarm : Alarm.DigitalAlarm;
END_VAR

(* One scan: Wanted members should run. *)
METHOD PROTECTED Coordinate
VAR_INPUT
    Wanted : INT;
END_VAR
VAR
    Index : INT;
    Count : INT;
    Active : INT;
    Running : INT;
    Available : INT;
    Pick : INT;
    Hours : LREAL;
    Best : LREAL;
END_VAR
    Members[1] := Member1;
    Members[2] := Member2;
    Members[3] := Member3;
    Members[4] := Member4;
    Count := 0;
    Active := 0;
    Running := 0;
    Available := 0;
    FOR Index := 1 TO 4 DO
        IF Members[Index] = NULL THEN
            Selected[Index] := FALSE;
        ELSE
            Count := Count + 1;
            (* A member that becomes unavailable is replaced. *)
            IF NOT Members[Index].IsAvailable() THEN
                Selected[Index] := FALSE;
            ELSE
                Available := Available + 1;
            END_IF;
            IF Members[Index].IsRunning() THEN
                Running := Running + 1;
            END_IF;
            IF Selected[Index] THEN
                Active := Active + 1;
            END_IF;
        END_IF;
    END_FOR;
    Target := LIMIT(0, Wanted, Count);

    (* One change at a time, StartDelay or StopDelay apart. *)
    SinceChange(IN := Changed, PT := T#24h);
    IF Active < Target AND (NOT Changed OR SinceChange.ET >= StartDelay) THEN
        Pick := 0;
        IF Preferred >= 1 AND Preferred <= 4 THEN
            IF Members[Preferred] <> NULL AND NOT Selected[Preferred] THEN
                IF Members[Preferred].IsAvailable() THEN
                    Pick := Preferred;
                END_IF;
            END_IF;
        END_IF;
        IF Pick = 0 THEN
            FOR Index := 1 TO 4 DO
                IF Members[Index] <> NULL AND NOT Selected[Index] THEN
                    IF Members[Index].IsAvailable() THEN
                        Hours := Members[Index].GetRunHours();
                        IF Pick = 0 OR Hours < Best THEN
                            Pick := Index;
                            Best := Hours;
                        END_IF;
                    END_IF;
                END_IF;
            END_FOR;
        END_IF;
        IF Pick > 0 THEN
            Selected[Pick] := TRUE;
            Changed := TRUE;
            SinceChange(IN := FALSE, PT := T#24h);
        END_IF;
    ELSIF Active > Target AND (NOT Changed OR SinceChange.ET >= StopDelay) THEN
        (* Stop the member that has run longest. *)
        Pick := 0;
        FOR Index := 1 TO 4 DO
            IF Selected[Index] THEN
                Hours := Members[Index].GetRunHours();
                IF Pick = 0 OR Hours > Best THEN
                    Pick := Index;
                    Best := Hours;
                END_IF;
            END_IF;
        END_FOR;
        IF Pick > 0 THEN
            Selected[Pick] := FALSE;
            Changed := TRUE;
            SinceChange(IN := FALSE, PT := T#24h);
        END_IF;
    END_IF;
    FOR Index := 1 TO 4 DO
        IF Members[Index] <> NULL THEN
            Members[Index].Demand(Run := Selected[Index]);
        END_IF;
    END_FOR;
    RunningCount := Running;
    AvailableCount := Available;
    ShortfallTimer(IN := Running < Target, PT := ShortfallDelay);
    Shortfall := ShortfallTimer.Q;
    ShortfallAlarm(Condition := Shortfall, Message := 'Not enough equipment available',
        Priority := AlarmPriority#High);
END_METHOD

METHOD PUBLIC GetAlarmCount : INT
    GetAlarmCount := 1;
END_METHOD

METHOD PUBLIC GetAlarm : REF_TO Alarm.Alarm
VAR_INPUT
    Index : INT;
END_VAR
    IF Index = 1 THEN
        GetAlarm := REF(ShortfallAlarm);
    ELSE
        GetAlarm := NULL;
    END_IF;
END_METHOD
END_FUNCTION_BLOCK

(* One member runs while Run is TRUE; a failed member is replaced by an available one. *)
FUNCTION_BLOCK FB_DutyStandbyGroup EXTENDS FB_Group
VAR_INPUT
    Run : BOOL;
END_VAR
    IF Run THEN
        Coordinate(Wanted := 1);
    ELSE
        Coordinate(Wanted := 0);
    END_IF;
END_FUNCTION_BLOCK

(* Required members run; the program decides how many. *)
FUNCTION_BLOCK FB_LeadLagGroup EXTENDS FB_Group
VAR_INPUT
    Required : INT;
END_VAR
    Coordinate(Wanted := Required);
END_FUNCTION_BLOCK

(* Demand in % of the group's equal stages, with hysteresis and minimum run and stop times. *)
FUNCTION_BLOCK FB_StagedGroup EXTENDS FB_Group
VAR_INPUT
    Demand : LREAL;
END_VAR
VAR PUBLIC RETAIN
    Hysteresis : LREAL := 5.0;
    MinRunTime : TIME := T#0s;
    MinStopTime : TIME := T#0s;
END_VAR
VAR NON_RETAIN
    Stages : INT;
    SinceStage : TON;
    Staged : BOOL;
END_VAR
VAR_TEMP
    Size : INT;
    StageSize : LREAL;
    Next : INT;
END_VAR
    Size := 0;
    IF Member1 <> NULL THEN Size := Size + 1; END_IF;
    IF Member2 <> NULL THEN Size := Size + 1; END_IF;
    IF Member3 <> NULL THEN Size := Size + 1; END_IF;
    IF Member4 <> NULL THEN Size := Size + 1; END_IF;
    Next := Stages;
    IF Size = 0 OR NOT F_Finite(Demand) OR Demand <= 0.0 THEN
        Next := 0;
    ELSE
        StageSize := 100.0 / INT_TO_LREAL(Size);
        WHILE Next < Size AND Demand > INT_TO_LREAL(Next) * StageSize DO
            Next := Next + 1;
        END_WHILE;
        WHILE Next > 1 AND Demand < INT_TO_LREAL(Next - 1) * StageSize - Hysteresis DO
            Next := Next - 1;
        END_WHILE;
    END_IF;
    SinceStage(IN := Staged, PT := T#24h);
    IF Next > Stages AND (NOT Staged OR SinceStage.ET >= MinStopTime) THEN
        Stages := Stages + 1;
        Staged := TRUE;
        SinceStage(IN := FALSE, PT := T#24h);
    ELSIF Next < Stages AND (NOT Staged OR SinceStage.ET >= MinRunTime) THEN
        Stages := Stages - 1;
        Staged := TRUE;
        SinceStage(IN := FALSE, PT := T#24h);
    END_IF;
    Coordinate(Wanted := Stages);
END_FUNCTION_BLOCK

END_NAMESPACE

(* ---- heater.st ---- *)
(* An electric heater (specification trust-plant-library §6.3): run control from FB_RunDevice for
   the main contactor, with the over-temperature switch as its trip, plus a power demand. A heater
   starts at 0 %: the operator's power is 0 % after a restart and after every stop. *)
NAMESPACE Plant

FUNCTION_BLOCK FB_Heater EXTENDS FB_RunDevice IMPLEMENTS IPowerDevice, IControlledDevice
VAR_INPUT
    (* The program's power in %, followed in Auto while running. *)
    AutoPower : LREAL;
END_VAR
VAR_OUTPUT NON_RETAIN
    (* The power in % for a thyristor controller. *)
    PowerOutput : LREAL;
    (* The same power, time-proportioned over PulsePeriod, for a solid-state relay. *)
    PulseOutput : BOOL;
    (* The operator's power in %. *)
    ManualPower : LREAL;
END_VAR
VAR PUBLIC RETAIN
    MaxPower : LREAL := 100.0;
    PulsePeriod : TIME := T#10s;
END_VAR
VAR NON_RETAIN
    WasCommanded : BOOL;
    Phase : TIME;
END_VAR
    ExecuteRun();
    ExecutePower();

METHOD PROTECTED ExecutePower
VAR
    High : LREAL;
    Wanted : LREAL;
    Period : LREAL;
END_VAR
    High := MAX(MaxPower, 0.0);
    IF RunCommand THEN
        IF Mode = E_Mode#Auto THEN
            Wanted := AutoPower;
            IF NOT F_Finite(Wanted) THEN
                Wanted := PowerOutput;
            END_IF;
            (* Bumpless: Manual continues at the power Auto had. *)
            ManualPower := LIMIT(0.0, Wanted, High);
        ELSE
            Wanted := ManualPower;
        END_IF;
        PowerOutput := LIMIT(0.0, Wanted, High);
    ELSE
        PowerOutput := 0.0;
        IF WasCommanded THEN
            ManualPower := 0.0;
        END_IF;
    END_IF;
    WasCommanded := RunCommand;

    (* Time proportioning: on for PowerOutput % of each period. *)
    Period := F_Seconds(PulsePeriod);
    IF RunCommand AND Period > 0.0 THEN
        Phase := Phase + Clock.Elapsed;
        IF Phase >= PulsePeriod THEN
            Phase := T#0s;
        END_IF;
        PulseOutput := F_Seconds(Phase) < Period * PowerOutput / 100.0;
    ELSE
        Phase := T#0s;
        PulseOutput := FALSE;
    END_IF;
END_METHOD

(* Accepted in Manual, also while stopped, so a power can be chosen before the start. *)
METHOD PUBLIC SetPower : BOOL
VAR_INPUT
    Value : LREAL;
END_VAR
    SetPower := AcceptsCommands() AND F_Finite(Value);
    IF SetPower THEN
        ManualPower := LIMIT(0.0, Value, MAX(MaxPower, 0.0));
    END_IF;
END_METHOD

(* The heater follows its Auto power while in Auto and running (§6.3); a controller that drives
   it tracks PowerOutput otherwise (§8.1). *)
METHOD PUBLIC FollowsAuto : BOOL
    FollowsAuto := Mode = E_Mode#Auto AND RunCommand;
END_METHOD

METHOD PUBLIC GetActualValue : LREAL
    GetActualValue := PowerOutput;
END_METHOD

END_FUNCTION_BLOCK

END_NAMESPACE

(* ---- managers.st ---- *)
(* Managers by composition (specification trust-plant-library §9.3, §9.4): the program names the
   blocks a manager covers in its call. Nothing registers. The HMI alarm list needs no manager:
   the runtime lists every alarm by itself. *)
NAMESPACE Plant

(* A summary of the alarms of up to sixteen blocks, for a horn or an area acknowledgement. *)
FUNCTION_BLOCK FB_AlarmManager IMPLEMENTS IAlarmManager
VAR_INPUT
    Source1 : IAlarmSource;
    Source2 : IAlarmSource;
    Source3 : IAlarmSource;
    Source4 : IAlarmSource;
    Source5 : IAlarmSource;
    Source6 : IAlarmSource;
    Source7 : IAlarmSource;
    Source8 : IAlarmSource;
    Source9 : IAlarmSource;
    Source10 : IAlarmSource;
    Source11 : IAlarmSource;
    Source12 : IAlarmSource;
    Source13 : IAlarmSource;
    Source14 : IAlarmSource;
    Source15 : IAlarmSource;
    Source16 : IAlarmSource;
END_VAR
VAR_OUTPUT NON_RETAIN
    ActiveCount : INT;
    UnacknowledgedCount : INT;
    (* TRUE from a new unacknowledged alarm until Silence or AcknowledgeAll. *)
    Horn : BOOL;
END_VAR
VAR NON_RETAIN
    Sources : ARRAY[1..16] OF IAlarmSource;
    Raised : ULINT;
    Primed : BOOL;
END_VAR
VAR_TEMP
    Index : INT;
    Item : INT;
    Total : ULINT;
    Entry : REF_TO Alarm.Alarm;
END_VAR
    Collect();
    ActiveCount := 0;
    UnacknowledgedCount := 0;
    Total := 0;
    FOR Index := 1 TO 16 DO
        IF Sources[Index] <> NULL THEN
            FOR Item := 1 TO Sources[Index].GetAlarmCount() DO
                Entry := Sources[Index].GetAlarm(Index := Item);
                IF Entry <> NULL THEN
                    (* A suppressed, shelved or out-of-service alarm is not counted (ISA-18.2). *)
                    IF Entry^.Active AND NOT (Entry^.SuppressedByDesign OR Entry^.Shelved OR Entry^.OutOfService) THEN
                        ActiveCount := ActiveCount + 1;
                    END_IF;
                    IF Entry^.Unacknowledged THEN
                        UnacknowledgedCount := UnacknowledgedCount + 1;
                    END_IF;
                    Total := Total + Entry^.AnnunciationCount;
                END_IF;
            END_FOR;
        END_IF;
    END_FOR;
    IF Primed AND Total > Raised THEN
        Horn := TRUE;
    END_IF;
    Raised := Total;
    Primed := TRUE;

METHOD PROTECTED Collect
    Sources[1] := Source1;
    Sources[2] := Source2;
    Sources[3] := Source3;
    Sources[4] := Source4;
    Sources[5] := Source5;
    Sources[6] := Source6;
    Sources[7] := Source7;
    Sources[8] := Source8;
    Sources[9] := Source9;
    Sources[10] := Source10;
    Sources[11] := Source11;
    Sources[12] := Source12;
    Sources[13] := Source13;
    Sources[14] := Source14;
    Sources[15] := Source15;
    Sources[16] := Source16;
END_METHOD

(* Acknowledges the alarms present now; an alarm raised later stays unacknowledged. *)
METHOD PUBLIC AcknowledgeAll : BOOL
VAR
    Index : INT;
    Item : INT;
    Entry : REF_TO Alarm.Alarm;
END_VAR
    Collect();
    FOR Index := 1 TO 16 DO
        IF Sources[Index] <> NULL THEN
            FOR Item := 1 TO Sources[Index].GetAlarmCount() DO
                Entry := Sources[Index].GetAlarm(Index := Item);
                IF Entry <> NULL THEN
                    Entry^.Acknowledge();
                END_IF;
            END_FOR;
        END_IF;
    END_FOR;
    Horn := FALSE;
    AcknowledgeAll := TRUE;
END_METHOD

METHOD PUBLIC Silence : BOOL
    Horn := FALSE;
    Silence := TRUE;
END_METHOD
END_FUNCTION_BLOCK

(* An overview of up to eight sequences; the program still executes each one. *)
FUNCTION_BLOCK FB_SequenceManager IMPLEMENTS ISequenceManager
VAR_INPUT
    Sequence1 : ISequence;
    Sequence2 : ISequence;
    Sequence3 : ISequence;
    Sequence4 : ISequence;
    Sequence5 : ISequence;
    Sequence6 : ISequence;
    Sequence7 : ISequence;
    Sequence8 : ISequence;
END_VAR
VAR_OUTPUT NON_RETAIN
    RunningCount : INT;
    HeldCount : INT;
    FailedCount : INT;
END_VAR
VAR NON_RETAIN
    Sequences : ARRAY[1..8] OF ISequence;
END_VAR
VAR_TEMP
    Index : INT;
    State : E_SequenceState;
END_VAR
    Collect();
    RunningCount := 0;
    HeldCount := 0;
    FailedCount := 0;
    FOR Index := 1 TO 8 DO
        IF Sequences[Index] <> NULL THEN
            State := Sequences[Index].GetState();
            IF State = E_SequenceState#Running OR State = E_SequenceState#Stopping THEN
                RunningCount := RunningCount + 1;
            ELSIF State = E_SequenceState#Held THEN
                HeldCount := HeldCount + 1;
            ELSIF State = E_SequenceState#Failed THEN
                FailedCount := FailedCount + 1;
            END_IF;
        END_IF;
    END_FOR;

METHOD PROTECTED Collect
    Sequences[1] := Sequence1;
    Sequences[2] := Sequence2;
    Sequences[3] := Sequence3;
    Sequences[4] := Sequence4;
    Sequences[5] := Sequence5;
    Sequences[6] := Sequence6;
    Sequences[7] := Sequence7;
    Sequences[8] := Sequence8;
END_METHOD

METHOD PUBLIC StopAll : BOOL
VAR
    Index : INT;
    Accepted : BOOL;
END_VAR
    Collect();
    StopAll := FALSE;
    FOR Index := 1 TO 8 DO
        IF Sequences[Index] <> NULL THEN
            Accepted := Sequences[Index].Stop();
            StopAll := StopAll OR Accepted;
        END_IF;
    END_FOR;
END_METHOD

METHOD PUBLIC AbortAll : BOOL
VAR
    Index : INT;
    Accepted : BOOL;
END_VAR
    Collect();
    AbortAll := FALSE;
    FOR Index := 1 TO 8 DO
        IF Sequences[Index] <> NULL THEN
            Accepted := Sequences[Index].Abort();
            AbortAll := AbortAll OR Accepted;
        END_IF;
    END_FOR;
END_METHOD
END_FUNCTION_BLOCK

END_NAMESPACE

(* ---- motor.st ---- *)
(* Run devices (specification trust-plant-library §6.1): one implementation of run control,
   feedback supervision, protection trips, counters and service, shared by the motor family, the
   variable-speed motors and the heater. *)
NAMESPACE Plant
USING Alarm;

FUNCTION_BLOCK ABSTRACT FB_RunDevice EXTENDS FB_Device IMPLEMENTS IDutyMember, IServiceable, IAlarmSource
VAR_INPUT
    (* The program's run demand, followed in Auto. *)
    AutoRun : BOOL;
    (* The run contact; ignored without HasFeedback. *)
    RunningFeedback : BOOL;
    (* A protection trip such as an overload relay: stops the device and latches. *)
    Trip : BOOL;
    HasFeedback : BOOL := TRUE;
END_VAR
VAR_OUTPUT NON_RETAIN
    (* The contactor output. *)
    RunCommand : BOOL;
    Running : BOOL;
    FailedToStart : BOOL;
    FailedToStop : BOOL;
    Tripped : BOOL;
    ServiceDue : BOOL;
END_VAR
VAR_OUTPUT RETAIN
    Starts : UDINT;
    RunHours : LREAL;
    HoursSinceService : LREAL;
END_VAR
VAR PUBLIC RETAIN
    StartTimeout : TIME := T#5s;
    StopTimeout : TIME := T#5s;
    (* Hours of running between services; 0 for none. *)
    ServiceInterval : LREAL := 4000.0;
END_VAR
VAR NON_RETAIN
    ManualRun : BOOL;
    GroupRun : BOOL;
    WasRunning : BOOL;
    StartWatch : TON;
    StopWatch : TON;
    Clock : FB_ScanClock;
    TripAlarm : Alarm.DigitalAlarm;
    FailedToStartAlarm : Alarm.DigitalAlarm;
    FailedToStopAlarm : Alarm.DigitalAlarm;
END_VAR

(* One scan of run control. A concrete block calls it from its body. *)
METHOD PROTECTED ExecuteRun
VAR
    Wanted : BOOL;
    Supervised : BOOL;
    Hours : LREAL;
END_VAR
    Clock();
    Supervised := Mode <> E_Mode#OutOfService;
    IF TakeReset() THEN
        IF NOT Trip THEN
            Tripped := FALSE;
        END_IF;
        FailedToStart := FALSE;
        FailedToStop := FALSE;
        StartWatch(IN := FALSE);
        StopWatch(IN := FALSE);
    END_IF;
    IF Supervised AND Trip THEN
        Tripped := TRUE;
    END_IF;
    Fault := Tripped OR FailedToStart OR FailedToStop;

    (* Who commands it (§3.2). *)
    CASE Mode OF
        E_Mode#Auto:
            Wanted := AutoRun OR GroupRun;
        E_Mode#Manual:
            Wanted := ManualRun;
    ELSE
        Wanted := FALSE;
    END_CASE;
    (* A start needs the permissive; a running device keeps running without it (§4.1). *)
    IF Wanted AND NOT RunCommand AND NOT MayStart() THEN
        Wanted := FALSE;
    END_IF;
    IF HeldSafe() THEN
        Wanted := FALSE;
    END_IF;
    RunCommand := Wanted;

    (* Feedback supervision, whoever commanded the device (§4.4). *)
    IF HasFeedback THEN
        Running := RunningFeedback;
    ELSE
        Running := RunCommand;
    END_IF;
    StartWatch(IN := Supervised AND HasFeedback AND RunCommand AND NOT RunningFeedback, PT := StartTimeout);
    StopWatch(IN := Supervised AND HasFeedback AND NOT RunCommand AND RunningFeedback, PT := StopTimeout);
    IF StartWatch.Q THEN
        FailedToStart := TRUE;
    END_IF;
    IF StopWatch.Q THEN
        FailedToStop := TRUE;
    END_IF;
    IF FailedToStart OR FailedToStop THEN
        Fault := TRUE;
        RunCommand := FALSE;
    END_IF;
    IF Tripped THEN
        FaultText := 'Protection trip: reset after the cause is cleared';
    ELSIF FailedToStart THEN
        FaultText := 'Failed to start: reset to try again';
    ELSIF FailedToStop THEN
        FaultText := 'Failed to stop: check the contactor, then reset';
    ELSE
        FaultText := '';
    END_IF;

    (* Bumpless (§3.4): Manual continues from the present command; any stop clears it. *)
    ManualRun := RunCommand;

    (* Alarms, suppressed by design only out of service (§4.5). *)
    TripAlarm(Condition := Tripped, Suppressed := NOT Supervised,
        Message := 'Protection trip', Priority := AlarmPriority#High);
    FailedToStartAlarm(Condition := FailedToStart, Suppressed := NOT Supervised,
        Message := 'Failed to start', Priority := AlarmPriority#Medium);
    FailedToStopAlarm(Condition := FailedToStop, Suppressed := NOT Supervised,
        Message := 'Failed to stop', Priority := AlarmPriority#High);

    (* Counters stand still out of service (§4.7). *)
    IF Supervised THEN
        IF Running AND NOT WasRunning AND Starts < UDINT#4294967295 THEN
            Starts := Starts + 1;
        END_IF;
        IF Running THEN
            Hours := Clock.Seconds / 3600.0;
            RunHours := RunHours + Hours;
            HoursSinceService := HoursSinceService + Hours;
        END_IF;
    END_IF;
    WasRunning := Running;
    ServiceDue := ServiceInterval > 0.0 AND HoursSinceService >= ServiceInterval;
    Publish();
END_METHOD

METHOD PUBLIC Start : BOOL
    Start := AcceptsStart();
    IF Start THEN
        ManualRun := TRUE;
    END_IF;
END_METHOD

METHOD PUBLIC Stop : BOOL
    Stop := AcceptsCommands();
    IF Stop THEN
        ManualRun := FALSE;
    END_IF;
END_METHOD

METHOD PUBLIC IsRunning : BOOL
    IsRunning := Running;
END_METHOD

(* A group may run it: in Auto, no fault, no interlock, and permitted or already running. *)
METHOD PUBLIC IsAvailable : BOOL
    IsAvailable := Mode = E_Mode#Auto AND NOT Fault AND NOT Interlock AND (Permissive OR RunCommand);
END_METHOD

(* A group's run demand, followed in Auto like AutoRun (§9.2). *)
METHOD PUBLIC Demand
VAR_INPUT
    Run : BOOL;
END_VAR
    GroupRun := Run;
END_METHOD

METHOD PUBLIC GetRunHours : LREAL
    GetRunHours := RunHours;
END_METHOD

METHOD PUBLIC ServiceDone : BOOL
    HoursSinceService := 0.0;
    ServiceDue := FALSE;
    ServiceDone := TRUE;
END_METHOD

METHOD PUBLIC GetAlarmCount : INT
    GetAlarmCount := 3;
END_METHOD

METHOD PUBLIC GetAlarm : REF_TO Alarm.Alarm
VAR_INPUT
    Index : INT;
END_VAR
    CASE Index OF
        1: GetAlarm := REF(TripAlarm);
        2: GetAlarm := REF(FailedToStartAlarm);
        3: GetAlarm := REF(FailedToStopAlarm);
    ELSE
        GetAlarm := NULL;
    END_CASE;
END_METHOD
END_FUNCTION_BLOCK

(* A fixed-speed motor. *)
FUNCTION_BLOCK FB_Motor EXTENDS FB_RunDevice
    ExecuteRun();
END_FUNCTION_BLOCK

(* The family below differs only in name and symbol; no process assumptions. *)
FUNCTION_BLOCK FB_Pump EXTENDS FB_Motor
    ExecuteRun();
END_FUNCTION_BLOCK

FUNCTION_BLOCK FB_Fan EXTENDS FB_Motor
    ExecuteRun();
END_FUNCTION_BLOCK

FUNCTION_BLOCK FB_Blower EXTENDS FB_Motor
    ExecuteRun();
END_FUNCTION_BLOCK

FUNCTION_BLOCK FB_Agitator EXTENDS FB_Motor
    ExecuteRun();
END_FUNCTION_BLOCK

FUNCTION_BLOCK FB_Conveyor EXTENDS FB_Motor
    ExecuteRun();
END_FUNCTION_BLOCK

END_NAMESPACE

(* ---- motor_valve.st ---- *)
(* A motor-operated valve (specification trust-plant-library §6.7). It has no spring: the motor
   drives it to an end limit and stops there, the operator may stop it in between, and its safe
   state stops it in place. Every movement counts as a start. *)
NAMESPACE Plant
USING Alarm;

FUNCTION_BLOCK FB_MotorValve EXTENDS FB_Device IMPLEMENTS IOpenCloseDevice, ITravelStop, IAlarmSource
VAR_INPUT
    (* The program's position, followed in Auto: TRUE open, FALSE closed. *)
    AutoOpen : BOOL;
    OpenLimit : BOOL;
    ClosedLimit : BOOL;
    (* The actuator's torque switch and the motor's overload relay; each latches. *)
    TorqueTrip : BOOL;
    Trip : BOOL;
END_VAR
VAR_OUTPUT NON_RETAIN
    OpenCommand : BOOL;
    CloseCommand : BOOL;
    Opened : BOOL;
    Closed : BOOL;
    Moving : BOOL;
    FailedToOpen : BOOL;
    FailedToClose : BOOL;
    FeedbackConflict : BOOL;
    Tripped : BOOL;
END_VAR
VAR_OUTPUT RETAIN
    Operations : UDINT;
END_VAR
VAR PUBLIC RETAIN
    TravelTimeout : TIME := T#60s;
END_VAR
VAR NON_RETAIN
    (* 0 stopped in place, 1 open, 2 closed: the target now and the operator's choice. *)
    Target : INT;
    ManualTarget : INT;
    WasOpened : BOOL;
    WasClosed : BOOL;
    Primed : BOOL;
    TravelWatch : TON;
    ConflictWatch : TON;
    TripAlarm : Alarm.DigitalAlarm;
    FailedToOpenAlarm : Alarm.DigitalAlarm;
    FailedToCloseAlarm : Alarm.DigitalAlarm;
END_VAR
    ExecuteTravel();

METHOD PROTECTED ExecuteTravel
VAR
    Wanted : INT;
    Supervised : BOOL;
    WasMoving : BOOL;
END_VAR
    Supervised := Mode <> E_Mode#OutOfService;
    IF TakeReset() THEN
        IF NOT Trip AND NOT TorqueTrip THEN
            Tripped := FALSE;
        END_IF;
        FailedToOpen := FALSE;
        FailedToClose := FALSE;
        FeedbackConflict := FALSE;
        TravelWatch(IN := FALSE);
        ConflictWatch(IN := FALSE);
    END_IF;
    IF Supervised AND (Trip OR TorqueTrip) THEN
        Tripped := TRUE;
    END_IF;
    Fault := Tripped OR FailedToOpen OR FailedToClose OR FeedbackConflict;

    CASE Mode OF
        E_Mode#Auto:
            IF AutoOpen THEN
                Wanted := 1;
            ELSE
                Wanted := 2;
            END_IF;
        E_Mode#Manual:
            Wanted := ManualTarget;
    ELSE
        Wanted := 0;
    END_CASE;
    WasMoving := OpenCommand OR CloseCommand;
    IF Wanted <> 0 AND Wanted <> Target AND NOT MayStart() THEN
        Wanted := 0;
    END_IF;
    IF HeldSafe() THEN
        Wanted := 0;
    END_IF;
    Target := Wanted;

    (* Drive towards the target until its limit, never both ways. *)
    OpenCommand := Target = 1 AND NOT OpenLimit;
    CloseCommand := Target = 2 AND NOT ClosedLimit;

    TravelWatch(IN := Supervised AND (OpenCommand OR CloseCommand), PT := TravelTimeout);
    IF TravelWatch.Q THEN
        IF OpenCommand THEN
            FailedToOpen := TRUE;
        ELSE
            FailedToClose := TRUE;
        END_IF;
    END_IF;
    ConflictWatch(IN := Supervised AND OpenLimit AND ClosedLimit, PT := T#1s);
    IF ConflictWatch.Q THEN
        FeedbackConflict := TRUE;
    END_IF;
    IF Tripped OR FailedToOpen OR FailedToClose OR FeedbackConflict THEN
        Fault := TRUE;
        Target := 0;
        OpenCommand := FALSE;
        CloseCommand := FALSE;
    END_IF;
    Opened := OpenLimit;
    Closed := ClosedLimit;
    Moving := OpenCommand OR CloseCommand;
    IF Tripped THEN
        FaultText := 'Motor or torque trip: reset after the cause is cleared';
    ELSIF FeedbackConflict THEN
        FaultText := 'Both limit switches active: check them, then reset';
    ELSIF FailedToOpen THEN
        FaultText := 'Did not open in time: reset to try again';
    ELSIF FailedToClose THEN
        FaultText := 'Did not close in time: reset to try again';
    ELSE
        FaultText := '';
    END_IF;

    (* Bumpless (§3.4); in Manual a refused or stopped movement leaves nothing pending. *)
    ManualTarget := Target;

    TripAlarm(Condition := Tripped, Suppressed := NOT Supervised,
        Message := 'Motor or torque trip', Priority := AlarmPriority#High);
    FailedToOpenAlarm(Condition := FailedToOpen, Suppressed := NOT Supervised,
        Message := 'Failed to open', Priority := AlarmPriority#Medium);
    FailedToCloseAlarm(Condition := FailedToClose OR FeedbackConflict, Suppressed := NOT Supervised,
        Message := 'Failed to close', Priority := AlarmPriority#Medium);
    IF Supervised AND Primed AND WasMoving
        AND ((OpenLimit AND NOT WasOpened) OR (ClosedLimit AND NOT WasClosed))
        AND Operations < UDINT#4294967295 THEN
        Operations := Operations + 1;
    END_IF;
    WasOpened := OpenLimit;
    WasClosed := ClosedLimit;
    Primed := TRUE;
    Publish();
END_METHOD

METHOD PUBLIC Open : BOOL
    Open := AcceptsStart();
    IF Open THEN
        ManualTarget := 1;
    END_IF;
END_METHOD

METHOD PUBLIC Close : BOOL
    Close := AcceptsStart();
    IF Close THEN
        ManualTarget := 2;
    END_IF;
END_METHOD

METHOD PUBLIC StopTravel : BOOL
    StopTravel := AcceptsCommands();
    IF StopTravel THEN
        ManualTarget := 0;
    END_IF;
END_METHOD

METHOD PUBLIC IsOpen : BOOL
    IsOpen := Opened;
END_METHOD

METHOD PUBLIC IsClosed : BOOL
    IsClosed := Closed;
END_METHOD

METHOD PUBLIC GetAlarmCount : INT
    GetAlarmCount := 3;
END_METHOD

METHOD PUBLIC GetAlarm : REF_TO Alarm.Alarm
VAR_INPUT
    Index : INT;
END_VAR
    CASE Index OF
        1: GetAlarm := REF(TripAlarm);
        2: GetAlarm := REF(FailedToOpenAlarm);
        3: GetAlarm := REF(FailedToCloseAlarm);
    ELSE
        GetAlarm := NULL;
    END_CASE;
END_METHOD
END_FUNCTION_BLOCK

END_NAMESPACE

(* ---- scale_and_tank.st ---- *)
(* The weigh scale and the tank (specification trust-plant-library §7.4, §7.5). *)
NAMESPACE Plant

(* An analog instrument with tare and stability. Tare is accepted only while the reading is
   stable and good. *)
FUNCTION_BLOCK FB_WeighScale EXTENDS FB_AnalogInput IMPLEMENTS ITare
VAR_OUTPUT NON_RETAIN
    Net : LREAL;
    Stable : BOOL;
END_VAR
VAR_OUTPUT RETAIN
    TareWeight : LREAL;
END_VAR
VAR PUBLIC RETAIN
    StableBand : LREAL := 0.5;
    StableTime : TIME := T#2s;
END_VAR
VAR NON_RETAIN
    Reference : LREAL;
    StableTimer : TON;
END_VAR
    Measure();
    Weigh();

METHOD PROTECTED Weigh
    IF Quality = E_Quality#Good AND ABS(Value - Reference) <= ABS(StableBand) THEN
        StableTimer(IN := TRUE, PT := StableTime);
    ELSE
        Reference := Value;
        StableTimer(IN := FALSE, PT := StableTime);
    END_IF;
    Stable := StableTimer.Q AND Quality = E_Quality#Good;
    Net := Value - TareWeight;
END_METHOD

METHOD PUBLIC Tare : BOOL
    Tare := Stable;
    IF Tare THEN
        TareWeight := Value;
        Net := 0.0;
    END_IF;
END_METHOD

METHOD PUBLIC ClearTare : BOOL
    TareWeight := 0.0;
    Net := Value;
    ClearTare := TRUE;
END_METHOD
END_FUNCTION_BLOCK

(* A tank shows the level of its level instrument, chosen by composition. It owns no filter and
   no alarms: the instrument owns them. *)
FUNCTION_BLOCK FB_Tank IMPLEMENTS IMeasurement
VAR_INPUT
    LevelInstrument : IMeasurement;
END_VAR
VAR PUBLIC RETAIN
    (* The level at 100 %. *)
    Height : LREAL := 100.0;
    (* The volume at Height; 0 when the volume is not shown. *)
    Capacity : LREAL := 0.0;
END_VAR
VAR_OUTPUT NON_RETAIN
    Level : LREAL;
    Percent : LREAL;
    Volume : LREAL;
    Quality : E_Quality := E_Quality#Bad;
END_VAR
    IF LevelInstrument = NULL THEN
        Quality := E_Quality#Bad;
    ELSE
        Level := LevelInstrument.GetValue();
        Quality := LevelInstrument.GetQuality();
    END_IF;
    IF Height > 0.0 THEN
        Percent := Level / Height * 100.0;
    ELSE
        Percent := 0.0;
    END_IF;
    IF Capacity > 0.0 THEN
        Volume := Capacity * Percent / 100.0;
    ELSE
        Volume := 0.0;
    END_IF;

METHOD PUBLIC GetValue : LREAL
    GetValue := Level;
END_METHOD

METHOD PUBLIC GetQuality : E_Quality
    GetQuality := Quality;
END_METHOD
END_FUNCTION_BLOCK

END_NAMESPACE

(* ---- sequence.st ---- *)
(* Sequences (specification trust-plant-library §9.4). FB_Sequence holds the lifecycle; an
   application sequence extends it, calls Execute from its body and writes its steps as a CASE on
   CurrentStep. Its outputs that command equipment are ordinary outputs wired to the devices' Auto inputs.
   Nothing is retained: after any restart a sequence is Idle. *)
NAMESPACE Plant

FUNCTION_BLOCK ABSTRACT FB_Sequence IMPLEMENTS ISequence
VAR_OUTPUT NON_RETAIN
    State : E_SequenceState;
    CurrentStep : INT;
    StepName : STRING[80];
    (* Time in the current step; it stands still while held. *)
    StepTime : TIME;
    (* What the sequence waits for, or why it failed. *)
    Message : STRING[120];
    (* The state in words, and which operator commands apply now. *)
    StateText : STRING[20] := 'Idle';
    CanStart : BOOL := TRUE;
    CanHold : BOOL;
    CanResume : BOOL;
    CanStop : BOOL;
    CanAbort : BOOL;
    CanReset : BOOL;
END_VAR
VAR NON_RETAIN
    Clock : FB_ScanClock;
END_VAR

(* The lifecycle of one scan; TRUE while Running, when the steps should advance. *)
METHOD PROTECTED Execute : BOOL
    Clock();
    IF State = E_SequenceState#Running OR State = E_SequenceState#Stopping THEN
        StepTime := StepTime + Clock.Elapsed;
    END_IF;
    Describe();
    Execute := State = E_SequenceState#Running;
END_METHOD

METHOD PROTECTED Describe
    CASE State OF
        E_SequenceState#Idle: StateText := 'Idle';
        E_SequenceState#Running: StateText := 'Running';
        E_SequenceState#Held: StateText := 'Held';
        E_SequenceState#Stopping: StateText := 'Stopping';
        E_SequenceState#Stopped: StateText := 'Stopped';
        E_SequenceState#Completed: StateText := 'Completed';
        E_SequenceState#Aborted: StateText := 'Aborted';
        E_SequenceState#Failed: StateText := 'Failed';
    END_CASE;
    CanStart := State = E_SequenceState#Idle;
    CanHold := State = E_SequenceState#Running;
    CanResume := State = E_SequenceState#Held;
    CanStop := State = E_SequenceState#Running OR State = E_SequenceState#Held;
    CanAbort := CanStop OR State = E_SequenceState#Stopping;
    CanReset := State = E_SequenceState#Stopped OR State = E_SequenceState#Completed
        OR State = E_SequenceState#Aborted OR State = E_SequenceState#Failed;
END_METHOD

(* Go to a step: its number and a name the operator reads. *)
METHOD PROTECTED GoTo
VAR_INPUT
    Number : INT;
    Name : STRING[80];
END_VAR
    CurrentStep := Number;
    StepName := Name;
    StepTime := T#0s;
    Message := '';
END_METHOD

(* Say what the step waits for. *)
METHOD PROTECTED Wait
VAR_INPUT
    Text : STRING[120];
END_VAR
    Message := Text;
END_METHOD

METHOD PROTECTED Complete
    IF State = E_SequenceState#Running THEN
        State := E_SequenceState#Completed;
        Message := '';
        Describe();
    END_IF;
END_METHOD

METHOD PROTECTED Fail
VAR_INPUT
    Text : STRING[120];
END_VAR
    IF State = E_SequenceState#Running OR State = E_SequenceState#Held
        OR State = E_SequenceState#Stopping THEN
        State := E_SequenceState#Failed;
        Message := Text;
        Describe();
    END_IF;
END_METHOD

(* The application's stop steps are done. *)
METHOD PROTECTED StopDone
    IF State = E_SequenceState#Stopping THEN
        State := E_SequenceState#Stopped;
        Describe();
    END_IF;
END_METHOD

(* Fails the sequence with Text when the current step has lasted longer than Limit. *)
METHOD PROTECTED StepTimeout : BOOL
VAR_INPUT
    Limit : TIME;
    Text : STRING[120];
END_VAR
    StepTimeout := State = E_SequenceState#Running AND StepTime > Limit;
    IF StepTimeout THEN
        Fail(Text := Text);
    END_IF;
END_METHOD

METHOD PUBLIC Start : BOOL
    Start := State = E_SequenceState#Idle;
    IF Start THEN
        State := E_SequenceState#Running;
        GoTo(Number := 0, Name := '');
        Describe();
    END_IF;
END_METHOD

METHOD PUBLIC Hold : BOOL
    Hold := State = E_SequenceState#Running;
    IF Hold THEN
        State := E_SequenceState#Held;
        Describe();
    END_IF;
END_METHOD

METHOD PUBLIC Resume : BOOL
    Resume := State = E_SequenceState#Held;
    IF Resume THEN
        State := E_SequenceState#Running;
        Describe();
    END_IF;
END_METHOD

METHOD PUBLIC Stop : BOOL
    Stop := State = E_SequenceState#Running OR State = E_SequenceState#Held;
    IF Stop THEN
        State := E_SequenceState#Stopping;
        Describe();
    END_IF;
END_METHOD

METHOD PUBLIC Abort : BOOL
    Abort := State = E_SequenceState#Running OR State = E_SequenceState#Held
        OR State = E_SequenceState#Stopping;
    IF Abort THEN
        State := E_SequenceState#Aborted;
        Message := 'Aborted by the operator';
        Describe();
    END_IF;
END_METHOD

METHOD PUBLIC Reset : BOOL
    Reset := State = E_SequenceState#Stopped OR State = E_SequenceState#Completed
        OR State = E_SequenceState#Aborted OR State = E_SequenceState#Failed;
    IF Reset THEN
        State := E_SequenceState#Idle;
        GoTo(Number := 0, Name := '');
        Describe();
    END_IF;
END_METHOD

METHOD PUBLIC GetState : E_SequenceState
    GetState := State;
END_METHOD
END_FUNCTION_BLOCK

END_NAMESPACE

(* ---- totals.st ---- *)
(* Accumulating instruments (specification trust-plant-library §7.3). *)
NAMESPACE Plant

(* Integrates a rate given per TotalPer; a bad or non-finite rate, and a rate at or below CutOff,
   is not counted. *)
FUNCTION_BLOCK FB_Totalizer IMPLEMENTS ITotal
VAR_INPUT
    (* The rate: an instrument by composition, else Rate and its quality. *)
    Measurement : IMeasurement;
    Rate : LREAL;
    RateGood : BOOL := TRUE;
END_VAR
VAR_OUTPUT RETAIN
    Total : LREAL;
END_VAR
VAR PUBLIC RETAIN
    TotalPer : TIME := T#1h;
    CutOff : LREAL := 0.0;
END_VAR
VAR NON_RETAIN
    Clock : FB_ScanClock;
END_VAR
VAR_TEMP
    Per : LREAL;
    Value : LREAL;
    Good : BOOL;
END_VAR
    Clock();
    IF Measurement <> NULL THEN
        Value := Measurement.GetValue();
        Good := Measurement.GetQuality() = E_Quality#Good;
    ELSE
        Value := Rate;
        Good := RateGood;
    END_IF;
    Per := F_Seconds(TotalPer);
    IF Good AND F_Finite(Value) AND Value > CutOff AND Per > 0.0 THEN
        Total := Total + Value * Clock.Seconds / Per;
    END_IF;

METHOD PUBLIC ResetTotal : BOOL
    Total := 0.0;
    ResetTotal := TRUE;
END_METHOD
END_FUNCTION_BLOCK

(* Counts rising edges of Pulse. A pulse that is already high after a restart is not counted. *)
FUNCTION_BLOCK FB_Counter IMPLEMENTS ICounter
VAR_INPUT
    Pulse : BOOL;
END_VAR
VAR_OUTPUT RETAIN
    Count : UDINT;
END_VAR
VAR_OUTPUT NON_RETAIN
    Done : BOOL;
END_VAR
VAR PUBLIC RETAIN
    (* Done at this count; 0 for none. *)
    Preset : UDINT := 0;
END_VAR
VAR NON_RETAIN
    Primed : BOOL;
    Previous : BOOL;
END_VAR
    IF Primed AND Pulse AND NOT Previous AND Count < UDINT#4294967295 THEN
        Count := Count + 1;
    END_IF;
    Previous := Pulse;
    Primed := TRUE;
    Done := Preset > 0 AND Count >= Preset;

METHOD PUBLIC ResetCount : BOOL
    Count := 0;
    Done := FALSE;
    ResetCount := TRUE;
END_METHOD
END_FUNCTION_BLOCK

END_NAMESPACE

(* ---- two_output_motor.st ---- *)
(* Motors with two exclusive run outputs (specification trust-plant-library §6.4, §6.5): the
   reversing motor (forward, reverse) and the two-speed motor (slow, fast). One implementation of
   the exclusive outputs, the transition delay, supervision, trips and counters; the concrete
   blocks name their own I/O. Direction or speed 0 is stopped, 1 is the first output, 2 the
   second. *)
NAMESPACE Plant
USING Alarm;

FUNCTION_BLOCK ABSTRACT FB_TwoOutputMotor EXTENDS FB_Device IMPLEMENTS IAlarmSource, IServiceable
VAR_INPUT
    Trip : BOOL;
    HasFeedback : BOOL := TRUE;
END_VAR
VAR_OUTPUT NON_RETAIN
    Running : BOOL;
    FailedToStart : BOOL;
    FailedToStop : BOOL;
    Tripped : BOOL;
    ServiceDue : BOOL;
END_VAR
VAR_OUTPUT RETAIN
    Starts : UDINT;
    RunHours : LREAL;
    HoursSinceService : LREAL;
END_VAR
VAR PUBLIC RETAIN
    StartTimeout : TIME := T#5s;
    StopTimeout : TIME := T#5s;
    (* Hours of running between services; 0 for none. *)
    ServiceInterval : LREAL := 4000.0;
END_VAR
VAR NON_RETAIN
    (* The output commanded now, the operator's choice, and the last running output. *)
    Commanded : INT;
    ManualWanted : INT;
    LastRun : INT;
    ActiveFirst : BOOL;
    ActiveSecond : BOOL;
    WasRunning : BOOL;
    Gap : TON;
    StartWatch : TON;
    StopWatch : TON;
    Clock : FB_ScanClock;
    TripAlarm : Alarm.DigitalAlarm;
    FailedToStartAlarm : Alarm.DigitalAlarm;
    FailedToStopAlarm : Alarm.DigitalAlarm;
END_VAR

(* One scan. AutoWanted is the program's choice; Delay is the transition time; with FullStop the
   motor must have stopped for Delay before the other output (reversing), else both outputs are
   simply dropped for Delay (changing speed). *)
METHOD PROTECTED ExecuteOutputs
VAR_INPUT
    AutoWanted : INT;
    FirstFeedback : BOOL;
    SecondFeedback : BOOL;
    Delay : TIME;
    FullStop : BOOL;
END_VAR
VAR
    Wanted : INT;
    Supervised : BOOL;
    Matching : BOOL;
    Hours : LREAL;
END_VAR
    Clock();
    Supervised := Mode <> E_Mode#OutOfService;
    IF TakeReset() THEN
        IF NOT Trip THEN
            Tripped := FALSE;
        END_IF;
        FailedToStart := FALSE;
        FailedToStop := FALSE;
        StartWatch(IN := FALSE);
        StopWatch(IN := FALSE);
    END_IF;
    IF Supervised AND Trip THEN
        Tripped := TRUE;
    END_IF;
    Fault := Tripped OR FailedToStart OR FailedToStop;

    CASE Mode OF
        E_Mode#Auto:
            Wanted := AutoWanted;
        E_Mode#Manual:
            Wanted := ManualWanted;
    ELSE
        Wanted := 0;
    END_CASE;
    IF Wanted < 0 OR Wanted > 2 THEN
        Wanted := 0;
    END_IF;
    (* A start, including one in the other direction or speed, needs the permissive. *)
    IF Wanted <> 0 AND Wanted <> Commanded AND NOT MayStart() THEN
        Wanted := 0;
    END_IF;
    IF HeldSafe() THEN
        Wanted := 0;
    END_IF;

    (* The transition: stop first, then the other output after the delay. *)
    IF Wanted = 0 THEN
        Commanded := 0;
    ELSIF Commanded <> 0 AND Commanded <> Wanted THEN
        Commanded := 0;
    END_IF;
    IF FullStop THEN
        Gap(IN := Commanded = 0 AND NOT Running, PT := Delay);
    ELSE
        Gap(IN := Commanded = 0, PT := Delay);
    END_IF;
    IF Commanded = 0 AND Wanted <> 0 THEN
        IF LastRun = 0 OR LastRun = Wanted OR Gap.Q THEN
            Commanded := Wanted;
        END_IF;
    END_IF;

    (* Feedback supervision (§4.4). *)
    IF HasFeedback THEN
        ActiveFirst := FirstFeedback;
        ActiveSecond := SecondFeedback;
    ELSE
        ActiveFirst := Commanded = 1;
        ActiveSecond := Commanded = 2;
    END_IF;
    Running := ActiveFirst OR ActiveSecond;
    Matching := (Commanded = 1 AND FirstFeedback AND NOT SecondFeedback)
        OR (Commanded = 2 AND SecondFeedback AND NOT FirstFeedback);
    StartWatch(IN := Supervised AND HasFeedback AND Commanded <> 0 AND NOT Matching, PT := StartTimeout);
    StopWatch(IN := Supervised AND HasFeedback AND Commanded = 0 AND Running, PT := StopTimeout);
    IF StartWatch.Q THEN
        FailedToStart := TRUE;
    END_IF;
    IF StopWatch.Q THEN
        FailedToStop := TRUE;
    END_IF;
    IF FailedToStart OR FailedToStop THEN
        Fault := TRUE;
        Commanded := 0;
        Wanted := 0;
    END_IF;
    IF Commanded <> 0 THEN
        LastRun := Commanded;
    END_IF;
    IF Tripped THEN
        FaultText := 'Protection trip: reset after the cause is cleared';
    ELSIF FailedToStart THEN
        FaultText := 'Failed to start: reset to try again';
    ELSIF FailedToStop THEN
        FaultText := 'Failed to stop: check the contactors, then reset';
    ELSE
        FaultText := '';
    END_IF;

    (* Bumpless (§3.4); a refused or stopped start leaves nothing pending in Manual. *)
    ManualWanted := Wanted;

    TripAlarm(Condition := Tripped, Suppressed := NOT Supervised,
        Message := 'Protection trip', Priority := AlarmPriority#High);
    FailedToStartAlarm(Condition := FailedToStart, Suppressed := NOT Supervised,
        Message := 'Failed to start', Priority := AlarmPriority#Medium);
    FailedToStopAlarm(Condition := FailedToStop, Suppressed := NOT Supervised,
        Message := 'Failed to stop', Priority := AlarmPriority#High);

    IF Supervised THEN
        IF Running AND NOT WasRunning AND Starts < UDINT#4294967295 THEN
            Starts := Starts + 1;
        END_IF;
        IF Running THEN
            Hours := Clock.Seconds / 3600.0;
            RunHours := RunHours + Hours;
            HoursSinceService := HoursSinceService + Hours;
        END_IF;
    END_IF;
    WasRunning := Running;
    ServiceDue := ServiceInterval > 0.0 AND HoursSinceService >= ServiceInterval;
    Publish();
END_METHOD

(* The service is done: the service count starts again; RunHours is unchanged (§4.7). *)
METHOD PUBLIC ServiceDone : BOOL
    HoursSinceService := 0.0;
    ServiceDue := FALSE;
    ServiceDone := TRUE;
END_METHOD

(* The operator's choice of output: accepted in Manual while nothing blocks a start. *)
METHOD PROTECTED RequestOutput : BOOL
VAR_INPUT
    Which : INT;
END_VAR
    RequestOutput := (Which = 1 OR Which = 2) AND AcceptsStart();
    IF RequestOutput THEN
        ManualWanted := Which;
    END_IF;
END_METHOD

METHOD PUBLIC Stop : BOOL
    Stop := AcceptsCommands();
    IF Stop THEN
        ManualWanted := 0;
    END_IF;
END_METHOD

METHOD PUBLIC GetAlarmCount : INT
    GetAlarmCount := 3;
END_METHOD

METHOD PUBLIC GetAlarm : REF_TO Alarm.Alarm
VAR_INPUT
    Index : INT;
END_VAR
    CASE Index OF
        1: GetAlarm := REF(TripAlarm);
        2: GetAlarm := REF(FailedToStartAlarm);
        3: GetAlarm := REF(FailedToStopAlarm);
    ELSE
        GetAlarm := NULL;
    END_CASE;
END_METHOD
END_FUNCTION_BLOCK

(* Forward and reverse. A change of direction stops the motor and waits ReversalDelay after it
   has stopped. Both Auto inputs TRUE means stop. *)
FUNCTION_BLOCK FB_ReversingMotor EXTENDS FB_TwoOutputMotor IMPLEMENTS IReversingDevice
VAR_INPUT
    AutoForward : BOOL;
    AutoReverse : BOOL;
    ForwardFeedback : BOOL;
    ReverseFeedback : BOOL;
END_VAR
VAR_OUTPUT NON_RETAIN
    ForwardCommand : BOOL;
    ReverseCommand : BOOL;
    Forward : BOOL;
    Reverse : BOOL;
END_VAR
VAR PUBLIC RETAIN
    ReversalDelay : TIME := T#2s;
END_VAR
VAR_TEMP
    Wanted : INT;
END_VAR
    IF AutoForward AND NOT AutoReverse THEN
        Wanted := 1;
    ELSIF AutoReverse AND NOT AutoForward THEN
        Wanted := 2;
    ELSE
        Wanted := 0;
    END_IF;
    ExecuteOutputs(AutoWanted := Wanted, FirstFeedback := ForwardFeedback,
        SecondFeedback := ReverseFeedback, Delay := ReversalDelay, FullStop := TRUE);
    ForwardCommand := Commanded = 1;
    ReverseCommand := Commanded = 2;
    Forward := ActiveFirst;
    Reverse := ActiveSecond;

METHOD PUBLIC StartForward : BOOL
    StartForward := RequestOutput(Which := 1);
END_METHOD

METHOD PUBLIC StartReverse : BOOL
    StartReverse := RequestOutput(Which := 2);
END_METHOD
END_FUNCTION_BLOCK

(* Slow and fast. Changing speed while running drops both outputs for ChangeoverDelay. *)
FUNCTION_BLOCK FB_TwoSpeedMotor EXTENDS FB_TwoOutputMotor IMPLEMENTS ITwoSpeedDevice
VAR_INPUT
    AutoRun : BOOL;
    AutoFast : BOOL;
    SlowFeedback : BOOL;
    FastFeedback : BOOL;
END_VAR
VAR_OUTPUT NON_RETAIN
    SlowCommand : BOOL;
    FastCommand : BOOL;
    Fast : BOOL;
END_VAR
VAR PUBLIC RETAIN
    ChangeoverDelay : TIME := T#1s;
END_VAR
VAR_TEMP
    Wanted : INT;
END_VAR
    IF NOT AutoRun THEN
        Wanted := 0;
    ELSIF AutoFast THEN
        Wanted := 2;
    ELSE
        Wanted := 1;
    END_IF;
    ExecuteOutputs(AutoWanted := Wanted, FirstFeedback := SlowFeedback,
        SecondFeedback := FastFeedback, Delay := ChangeoverDelay, FullStop := FALSE);
    SlowCommand := Commanded = 1;
    FastCommand := Commanded = 2;
    Fast := ActiveSecond;

METHOD PUBLIC StartSlow : BOOL
    StartSlow := RequestOutput(Which := 1);
END_METHOD

METHOD PUBLIC StartFast : BOOL
    StartFast := RequestOutput(Which := 2);
END_METHOD
END_FUNCTION_BLOCK

END_NAMESPACE

(* ---- valve.st ---- *)
(* On/off valves and dampers (specification trust-plant-library §6.6). The safe state is the fail
   position: the de-energised solenoid, closed or, with FailOpen, open. Moving away from the fail
   position counts as a start: it needs the permissive and is refused while blocked. *)
NAMESPACE Plant
USING Alarm;

FUNCTION_BLOCK FB_OnOffValve EXTENDS FB_Device IMPLEMENTS IOpenCloseDevice, IAlarmSource
VAR_INPUT
    (* The program's position, followed in Auto: TRUE open. *)
    AutoOpen : BOOL;
    OpenFeedback : BOOL;
    ClosedFeedback : BOOL;
    HasOpenFeedback : BOOL := TRUE;
    HasClosedFeedback : BOOL := TRUE;
    (* The valve opens when its solenoid loses power. *)
    FailOpen : BOOL;
END_VAR
VAR_OUTPUT NON_RETAIN
    (* The commanded position: TRUE open. *)
    OpenCommand : BOOL;
    (* The solenoid output: energised to leave the fail position. *)
    Solenoid : BOOL;
    Opened : BOOL;
    Closed : BOOL;
    Moving : BOOL;
    FailedToOpen : BOOL;
    FailedToClose : BOOL;
    FeedbackConflict : BOOL;
    (* The operator may open, or close, now. *)
    OpenPermit : BOOL;
    ClosePermit : BOOL;
END_VAR
VAR_OUTPUT RETAIN
    Operations : UDINT;
END_VAR
VAR PUBLIC RETAIN
    OpenTimeout : TIME := T#10s;
    CloseTimeout : TIME := T#10s;
END_VAR
VAR NON_RETAIN
    ManualOpen : BOOL;
    Initialized : BOOL;
    Watch : FB_EndPositionWatch;
    FailedToOpenAlarm : Alarm.DigitalAlarm;
    FailedToCloseAlarm : Alarm.DigitalAlarm;
    ConflictAlarm : Alarm.DigitalAlarm;
END_VAR
    ExecuteValve();

METHOD PROTECTED ExecuteValve
VAR
    Wanted : BOOL;
    Supervised : BOOL;
END_VAR
    (* After a restart a manually commanded valve is in its fail position (§4.8). *)
    IF NOT Initialized THEN
        ManualOpen := FailOpen;
        OpenCommand := FailOpen;
        Initialized := TRUE;
    END_IF;
    Supervised := Mode <> E_Mode#OutOfService;
    CASE Mode OF
        E_Mode#Auto:
            Wanted := AutoOpen;
        E_Mode#Manual:
            Wanted := ManualOpen;
    ELSE
        Wanted := FailOpen;
    END_CASE;
    IF Wanted <> FailOpen AND OpenCommand = FailOpen AND NOT MayStart() THEN
        Wanted := FailOpen;
    END_IF;
    IF HeldSafe() THEN
        Wanted := FailOpen;
    END_IF;
    OpenCommand := Wanted;

    Watch(Enable := Supervised, TowardsA := OpenCommand, AtA := OpenFeedback, AtB := ClosedFeedback,
        HasA := HasOpenFeedback, HasB := HasClosedFeedback, TimeoutA := OpenTimeout,
        TimeoutB := CloseTimeout, Clear := TakeReset());
    FailedToOpen := Watch.FailedA;
    FailedToClose := Watch.FailedB;
    FeedbackConflict := Watch.Conflict;
    Fault := FailedToOpen OR FailedToClose OR FeedbackConflict;
    IF Fault THEN
        OpenCommand := FailOpen;
    END_IF;
    Solenoid := OpenCommand XOR FailOpen;
    Opened := Watch.InA;
    Closed := Watch.InB;
    Moving := Watch.Moving;
    IF FeedbackConflict THEN
        FaultText := 'Both end switches active: check them, then reset';
    ELSIF FailedToOpen THEN
        FaultText := 'Failed to open: reset to try again';
    ELSIF FailedToClose THEN
        FaultText := 'Failed to close: reset to try again';
    ELSE
        FaultText := '';
    END_IF;

    (* Bumpless (§3.4). *)
    ManualOpen := OpenCommand;

    FailedToOpenAlarm(Condition := FailedToOpen, Suppressed := NOT Supervised,
        Message := 'Failed to open', Priority := AlarmPriority#Medium);
    FailedToCloseAlarm(Condition := FailedToClose, Suppressed := NOT Supervised,
        Message := 'Failed to close', Priority := AlarmPriority#Medium);
    ConflictAlarm(Condition := FeedbackConflict, Suppressed := NOT Supervised,
        Message := 'End switches conflict', Priority := AlarmPriority#Medium);
    IF Supervised AND Watch.Arrived AND Operations < UDINT#4294967295 THEN
        Operations := Operations + 1;
    END_IF;
    Publish();
    OpenPermit := Manual AND (FailOpen OR NOT Blocked);
    ClosePermit := Manual AND (NOT FailOpen OR NOT Blocked);
END_METHOD

METHOD PUBLIC Open : BOOL
    IF FailOpen THEN
        Open := AcceptsCommands();
    ELSE
        Open := AcceptsStart();
    END_IF;
    IF Open THEN
        ManualOpen := TRUE;
    END_IF;
END_METHOD

METHOD PUBLIC Close : BOOL
    IF FailOpen THEN
        Close := AcceptsStart();
    ELSE
        Close := AcceptsCommands();
    END_IF;
    IF Close THEN
        ManualOpen := FALSE;
    END_IF;
END_METHOD

METHOD PUBLIC IsOpen : BOOL
    IsOpen := Opened;
END_METHOD

METHOD PUBLIC IsClosed : BOOL
    IsClosed := Closed;
END_METHOD

METHOD PUBLIC GetAlarmCount : INT
    GetAlarmCount := 3;
END_METHOD

METHOD PUBLIC GetAlarm : REF_TO Alarm.Alarm
VAR_INPUT
    Index : INT;
END_VAR
    CASE Index OF
        1: GetAlarm := REF(FailedToOpenAlarm);
        2: GetAlarm := REF(FailedToCloseAlarm);
        3: GetAlarm := REF(ConflictAlarm);
    ELSE
        GetAlarm := NULL;
    END_CASE;
END_METHOD
END_FUNCTION_BLOCK

(* An on/off damper: the valve's behaviour with a damper's name and symbol. *)
FUNCTION_BLOCK FB_Damper EXTENDS FB_OnOffValve
    ExecuteValve();
END_FUNCTION_BLOCK

END_NAMESPACE
